// TIA Portal V18 export
FUNCTION "Interlock dos sinais linha" : Void   // FC9, LAD
{ S7_Optimized_Access := 'TRUE' }
// stored: SetENOAutomatically false
   VAR_TEMP
      SIGNAL_HELGE : Bool;
      SIGNAL_HELGE1 : Bool;
   END_VAR
   VAR_TEMP   // added for the SCL form of the ladder/FBD networks
      _w1 : Bool;
      _w2 : Bool;
      _w3 : Bool;
      _w4 : Bool;
   END_VAR
BEGIN

REGION Network 1: SCADA DESABILITADO
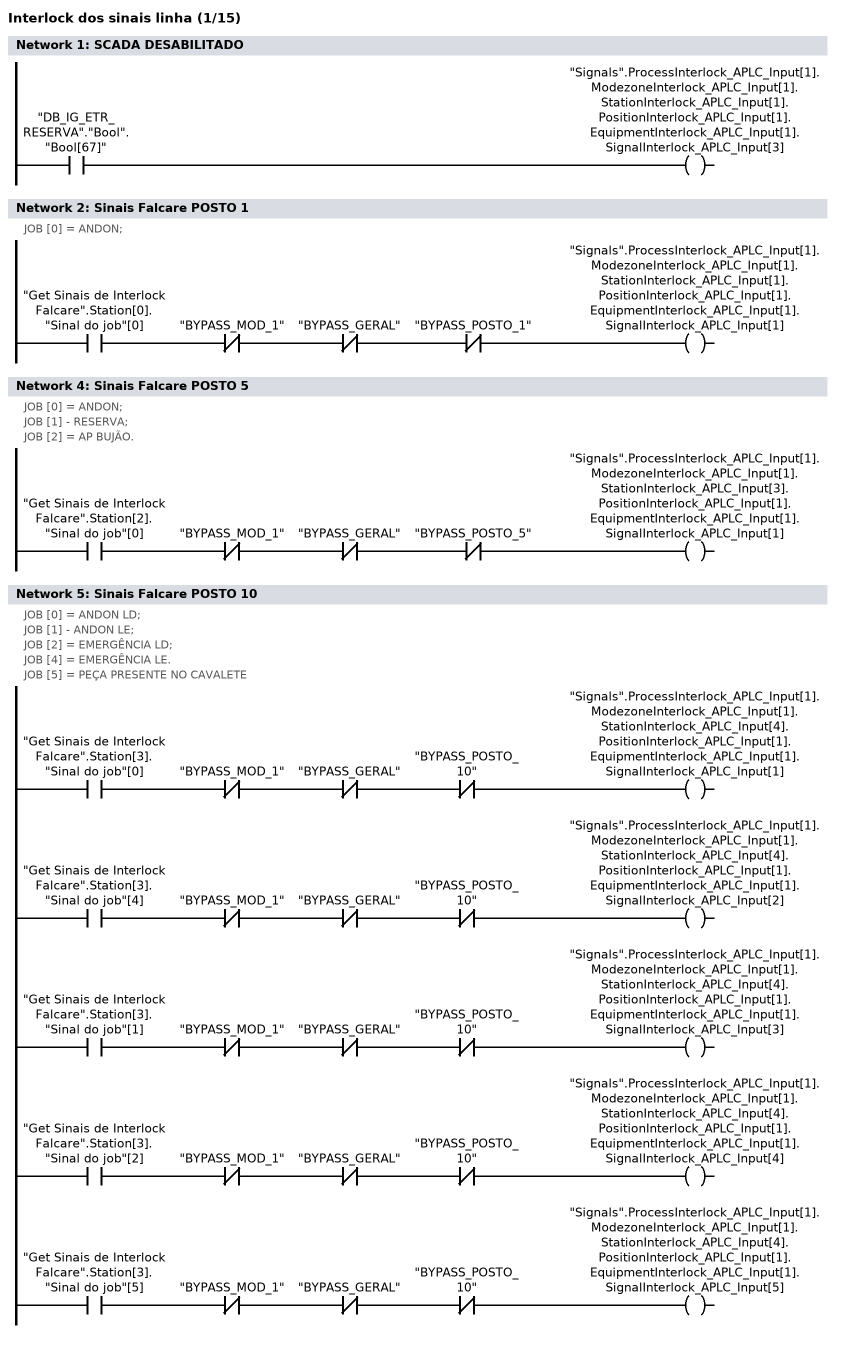
   RUNG wire#powerrail
      Contact( "DB_IG_ETR_RESERVA"."Bool"."Bool[67]" )
      Coil( "Signals".ProcessInterlock_APLC_Input[1].ModezoneInterlock_APLC_Input[1].StationInterlock_APLC_Input[1].PositionInterlock_APLC_Input[1].EquipmentInterlock_APLC_Input[1].SignalInterlock_APLC_Input[3] )
   END_RUNG
   // the same network as SCL:
   "Signals".ProcessInterlock_APLC_Input[1].ModezoneInterlock_APLC_Input[1].StationInterlock_APLC_Input[1].PositionInterlock_APLC_Input[1].EquipmentInterlock_APLC_Input[1].SignalInterlock_APLC_Input[3] := "DB_IG_ETR_RESERVA"."Bool"."Bool[67]";
END_REGION

REGION Network 2: Sinais Falcare POSTO 1
   // JOB [0] = ANDON;
   RUNG wire#powerrail
      Contact( "Get Sinais de Interlock Falcare".Station[0]."Sinal do job"[0] )
      I_Contact( "BYPASS_MOD_1" )
      I_Contact( "BYPASS_GERAL" )
      I_Contact( "BYPASS_POSTO_1" )
      Coil( "Signals".ProcessInterlock_APLC_Input[1].ModezoneInterlock_APLC_Input[1].StationInterlock_APLC_Input[1].PositionInterlock_APLC_Input[1].EquipmentInterlock_APLC_Input[1].SignalInterlock_APLC_Input[1] )
   END_RUNG
   // the same network as SCL:
   "Signals".ProcessInterlock_APLC_Input[1].ModezoneInterlock_APLC_Input[1].StationInterlock_APLC_Input[1].PositionInterlock_APLC_Input[1].EquipmentInterlock_APLC_Input[1].SignalInterlock_APLC_Input[1] := "Get Sinais de Interlock Falcare".Station[0]."Sinal do job"[0] AND NOT "BYPASS_MOD_1" AND NOT "BYPASS_GERAL" AND NOT "BYPASS_POSTO_1";
END_REGION

REGION Network 3: Sinais Falcare VIVERK
   // JOB [0] = ANDON;
   // JOB [1] - EMERGÊNCIA;
END_REGION

REGION Network 4: Sinais Falcare POSTO 5
   // JOB [0] = ANDON;
   // JOB [1] - RESERVA;
   // JOB [2] = AP BUJÃO.
   RUNG wire#powerrail
      Contact( "Get Sinais de Interlock Falcare".Station[2]."Sinal do job"[0] )
      I_Contact( "BYPASS_MOD_1" )
      I_Contact( "BYPASS_GERAL" )
      I_Contact( "BYPASS_POSTO_5" )
      Coil( "Signals".ProcessInterlock_APLC_Input[1].ModezoneInterlock_APLC_Input[1].StationInterlock_APLC_Input[3].PositionInterlock_APLC_Input[1].EquipmentInterlock_APLC_Input[1].SignalInterlock_APLC_Input[1] )
   END_RUNG
   // the same network as SCL:
   "Signals".ProcessInterlock_APLC_Input[1].ModezoneInterlock_APLC_Input[1].StationInterlock_APLC_Input[3].PositionInterlock_APLC_Input[1].EquipmentInterlock_APLC_Input[1].SignalInterlock_APLC_Input[1] := "Get Sinais de Interlock Falcare".Station[2]."Sinal do job"[0] AND NOT "BYPASS_MOD_1" AND NOT "BYPASS_GERAL" AND NOT "BYPASS_POSTO_5";
END_REGION

REGION Network 5: Sinais Falcare POSTO 10
   // JOB [0] = ANDON LD;
   // JOB [1] - ANDON LE;
   // JOB [2] = EMERGÊNCIA LD;
   // JOB [4] = EMERGÊNCIA LE.
   // JOB [5] = PEÇA PRESENTE NO CAVALETE
   RUNG wire#powerrail
      Contact( "Get Sinais de Interlock Falcare".Station[3]."Sinal do job"[0] )
      I_Contact( "BYPASS_MOD_1" )
      I_Contact( "BYPASS_GERAL" )
      I_Contact( "BYPASS_POSTO_10" )
      Coil( "Signals".ProcessInterlock_APLC_Input[1].ModezoneInterlock_APLC_Input[1].StationInterlock_APLC_Input[4].PositionInterlock_APLC_Input[1].EquipmentInterlock_APLC_Input[1].SignalInterlock_APLC_Input[1] )
   END_RUNG
   RUNG wire#powerrail
      Contact( "Get Sinais de Interlock Falcare".Station[3]."Sinal do job"[4] )
      I_Contact( "BYPASS_MOD_1" )
      I_Contact( "BYPASS_GERAL" )
      I_Contact( "BYPASS_POSTO_10" )
      Coil( "Signals".ProcessInterlock_APLC_Input[1].ModezoneInterlock_APLC_Input[1].StationInterlock_APLC_Input[4].PositionInterlock_APLC_Input[1].EquipmentInterlock_APLC_Input[1].SignalInterlock_APLC_Input[2] )
   END_RUNG
   RUNG wire#powerrail
      Contact( "Get Sinais de Interlock Falcare".Station[3]."Sinal do job"[1] )
      I_Contact( "BYPASS_MOD_1" )
      I_Contact( "BYPASS_GERAL" )
      I_Contact( "BYPASS_POSTO_10" )
      Coil( "Signals".ProcessInterlock_APLC_Input[1].ModezoneInterlock_APLC_Input[1].StationInterlock_APLC_Input[4].PositionInterlock_APLC_Input[1].EquipmentInterlock_APLC_Input[1].SignalInterlock_APLC_Input[3] )
   END_RUNG
   RUNG wire#powerrail
      Contact( "Get Sinais de Interlock Falcare".Station[3]."Sinal do job"[2] )
      I_Contact( "BYPASS_MOD_1" )
      I_Contact( "BYPASS_GERAL" )
      I_Contact( "BYPASS_POSTO_10" )
      Coil( "Signals".ProcessInterlock_APLC_Input[1].ModezoneInterlock_APLC_Input[1].StationInterlock_APLC_Input[4].PositionInterlock_APLC_Input[1].EquipmentInterlock_APLC_Input[1].SignalInterlock_APLC_Input[4] )
   END_RUNG
   RUNG wire#powerrail
      Contact( "Get Sinais de Interlock Falcare".Station[3]."Sinal do job"[5] )
      I_Contact( "BYPASS_MOD_1" )
      I_Contact( "BYPASS_GERAL" )
      I_Contact( "BYPASS_POSTO_10" )
      Coil( "Signals".ProcessInterlock_APLC_Input[1].ModezoneInterlock_APLC_Input[1].StationInterlock_APLC_Input[4].PositionInterlock_APLC_Input[1].EquipmentInterlock_APLC_Input[1].SignalInterlock_APLC_Input[5] )
   END_RUNG
   // the same network as SCL:
   "Signals".ProcessInterlock_APLC_Input[1].ModezoneInterlock_APLC_Input[1].StationInterlock_APLC_Input[4].PositionInterlock_APLC_Input[1].EquipmentInterlock_APLC_Input[1].SignalInterlock_APLC_Input[1] := "Get Sinais de Interlock Falcare".Station[3]."Sinal do job"[0] AND NOT "BYPASS_MOD_1" AND NOT "BYPASS_GERAL" AND NOT "BYPASS_POSTO_10";
   "Signals".ProcessInterlock_APLC_Input[1].ModezoneInterlock_APLC_Input[1].StationInterlock_APLC_Input[4].PositionInterlock_APLC_Input[1].EquipmentInterlock_APLC_Input[1].SignalInterlock_APLC_Input[2] := "Get Sinais de Interlock Falcare".Station[3]."Sinal do job"[4] AND NOT "BYPASS_MOD_1" AND NOT "BYPASS_GERAL" AND NOT "BYPASS_POSTO_10";
   "Signals".ProcessInterlock_APLC_Input[1].ModezoneInterlock_APLC_Input[1].StationInterlock_APLC_Input[4].PositionInterlock_APLC_Input[1].EquipmentInterlock_APLC_Input[1].SignalInterlock_APLC_Input[3] := "Get Sinais de Interlock Falcare".Station[3]."Sinal do job"[1] AND NOT "BYPASS_MOD_1" AND NOT "BYPASS_GERAL" AND NOT "BYPASS_POSTO_10";
   "Signals".ProcessInterlock_APLC_Input[1].ModezoneInterlock_APLC_Input[1].StationInterlock_APLC_Input[4].PositionInterlock_APLC_Input[1].EquipmentInterlock_APLC_Input[1].SignalInterlock_APLC_Input[4] := "Get Sinais de Interlock Falcare".Station[3]."Sinal do job"[2] AND NOT "BYPASS_MOD_1" AND NOT "BYPASS_GERAL" AND NOT "BYPASS_POSTO_10";
   "Signals".ProcessInterlock_APLC_Input[1].ModezoneInterlock_APLC_Input[1].StationInterlock_APLC_Input[4].PositionInterlock_APLC_Input[1].EquipmentInterlock_APLC_Input[1].SignalInterlock_APLC_Input[5] := "Get Sinais de Interlock Falcare".Station[3]."Sinal do job"[5] AND NOT "BYPASS_MOD_1" AND NOT "BYPASS_GERAL" AND NOT "BYPASS_POSTO_10";
END_REGION

REGION Network 6: Sinais Falcare POSTO 15
   // JOB [3] = AP TUBO RPX POSTO 15;
END_REGION

REGION Network 7: Sinais Falcare POSTO 20
   // JOB [0] = ANDON LD;
   // JOB [1] - EMERGÊNCIA LD;
   // JOB [2] = AP MOLA HARPA;
   // JOB [3] = SENSOR POSIÇÃO AP HARPA;
   // JOB [4] = AP TUBO LUBRIFICAÇÃO RPX I9.0
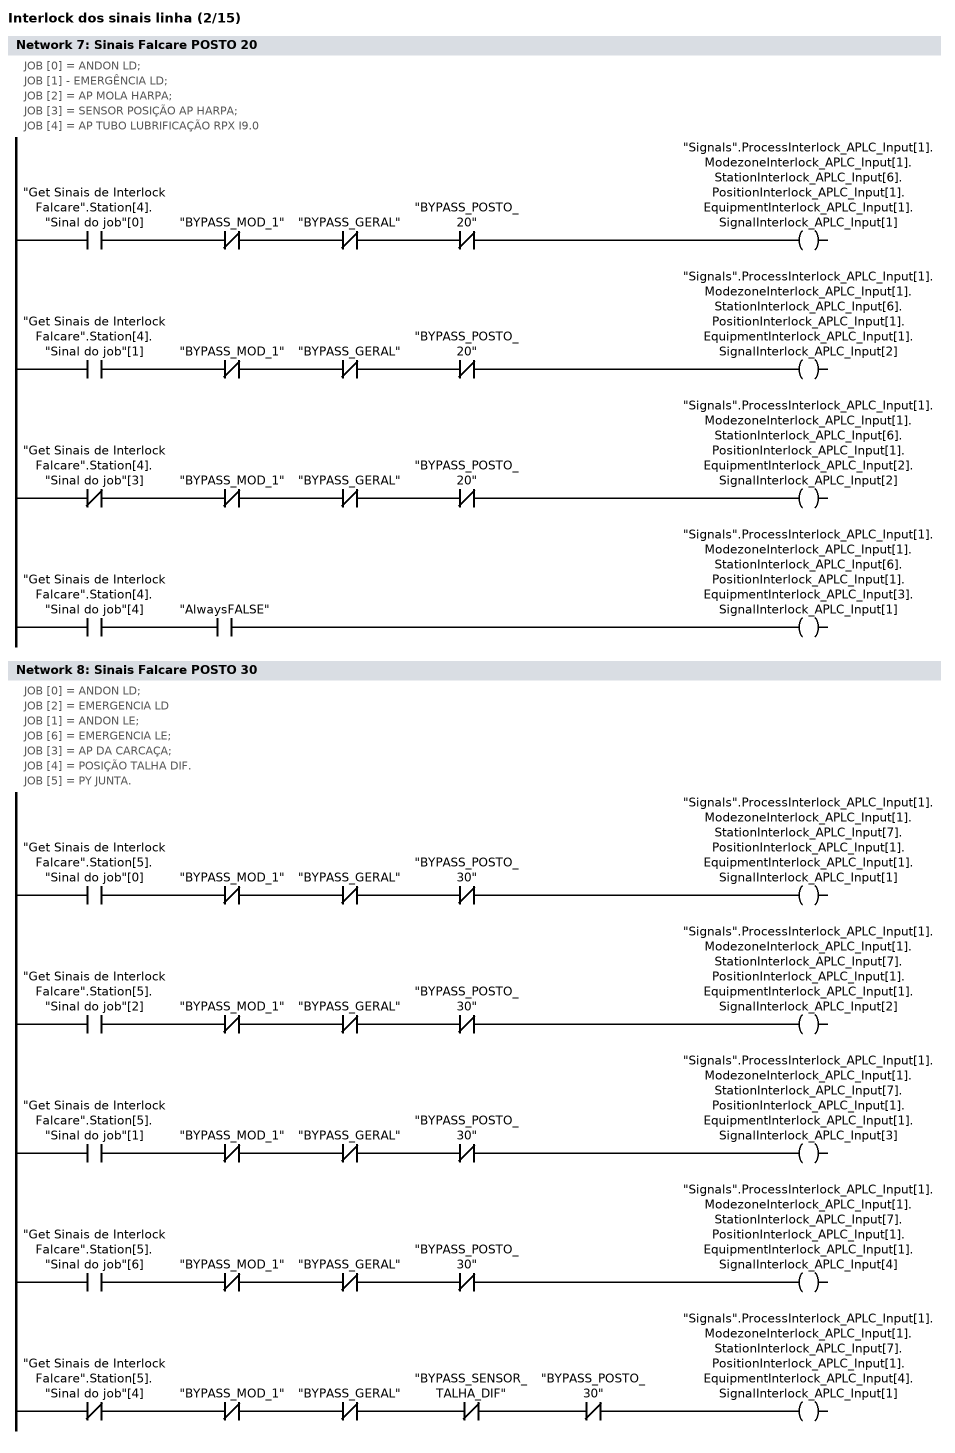
   RUNG wire#powerrail
      Contact( "Get Sinais de Interlock Falcare".Station[4]."Sinal do job"[0] )
      I_Contact( "BYPASS_MOD_1" )
      I_Contact( "BYPASS_GERAL" )
      I_Contact( "BYPASS_POSTO_20" )
      Coil( "Signals".ProcessInterlock_APLC_Input[1].ModezoneInterlock_APLC_Input[1].StationInterlock_APLC_Input[6].PositionInterlock_APLC_Input[1].EquipmentInterlock_APLC_Input[1].SignalInterlock_APLC_Input[1] )
   END_RUNG
   RUNG wire#powerrail
      Contact( "Get Sinais de Interlock Falcare".Station[4]."Sinal do job"[1] )
      I_Contact( "BYPASS_MOD_1" )
      I_Contact( "BYPASS_GERAL" )
      I_Contact( "BYPASS_POSTO_20" )
      Coil( "Signals".ProcessInterlock_APLC_Input[1].ModezoneInterlock_APLC_Input[1].StationInterlock_APLC_Input[6].PositionInterlock_APLC_Input[1].EquipmentInterlock_APLC_Input[1].SignalInterlock_APLC_Input[2] )
   END_RUNG
   RUNG wire#powerrail
      I_Contact( "Get Sinais de Interlock Falcare".Station[4]."Sinal do job"[3] )
      I_Contact( "BYPASS_MOD_1" )
      I_Contact( "BYPASS_GERAL" )
      I_Contact( "BYPASS_POSTO_20" )
      Coil( "Signals".ProcessInterlock_APLC_Input[1].ModezoneInterlock_APLC_Input[1].StationInterlock_APLC_Input[6].PositionInterlock_APLC_Input[1].EquipmentInterlock_APLC_Input[2].SignalInterlock_APLC_Input[2] )
   END_RUNG
   RUNG wire#powerrail
      Contact( "Get Sinais de Interlock Falcare".Station[4]."Sinal do job"[4] )
      Contact( "AlwaysFALSE" )
      Coil( "Signals".ProcessInterlock_APLC_Input[1].ModezoneInterlock_APLC_Input[1].StationInterlock_APLC_Input[6].PositionInterlock_APLC_Input[1].EquipmentInterlock_APLC_Input[3].SignalInterlock_APLC_Input[1] )
   END_RUNG
   // the same network as SCL:
   "Signals".ProcessInterlock_APLC_Input[1].ModezoneInterlock_APLC_Input[1].StationInterlock_APLC_Input[6].PositionInterlock_APLC_Input[1].EquipmentInterlock_APLC_Input[1].SignalInterlock_APLC_Input[1] := "Get Sinais de Interlock Falcare".Station[4]."Sinal do job"[0] AND NOT "BYPASS_MOD_1" AND NOT "BYPASS_GERAL" AND NOT "BYPASS_POSTO_20";
   "Signals".ProcessInterlock_APLC_Input[1].ModezoneInterlock_APLC_Input[1].StationInterlock_APLC_Input[6].PositionInterlock_APLC_Input[1].EquipmentInterlock_APLC_Input[1].SignalInterlock_APLC_Input[2] := "Get Sinais de Interlock Falcare".Station[4]."Sinal do job"[1] AND NOT "BYPASS_MOD_1" AND NOT "BYPASS_GERAL" AND NOT "BYPASS_POSTO_20";
   "Signals".ProcessInterlock_APLC_Input[1].ModezoneInterlock_APLC_Input[1].StationInterlock_APLC_Input[6].PositionInterlock_APLC_Input[1].EquipmentInterlock_APLC_Input[2].SignalInterlock_APLC_Input[2] := NOT "Get Sinais de Interlock Falcare".Station[4]."Sinal do job"[3] AND NOT "BYPASS_MOD_1" AND NOT "BYPASS_GERAL" AND NOT "BYPASS_POSTO_20";
   "Signals".ProcessInterlock_APLC_Input[1].ModezoneInterlock_APLC_Input[1].StationInterlock_APLC_Input[6].PositionInterlock_APLC_Input[1].EquipmentInterlock_APLC_Input[3].SignalInterlock_APLC_Input[1] := "Get Sinais de Interlock Falcare".Station[4]."Sinal do job"[4] AND "AlwaysFALSE";
END_REGION

REGION Network 8: Sinais Falcare POSTO 30
   // JOB [0] = ANDON LD;
   // JOB [2] = EMERGENCIA LD
   // JOB [1] = ANDON LE;
   // JOB [6] = EMERGENCIA LE;
   // JOB [3] = AP DA CARCAÇA;
   // JOB [4] = POSIÇÃO TALHA DIF.
   // JOB [5] = PY JUNTA.
   RUNG wire#powerrail
      Contact( "Get Sinais de Interlock Falcare".Station[5]."Sinal do job"[0] )
      I_Contact( "BYPASS_MOD_1" )
      I_Contact( "BYPASS_GERAL" )
      I_Contact( "BYPASS_POSTO_30" )
      Coil( "Signals".ProcessInterlock_APLC_Input[1].ModezoneInterlock_APLC_Input[1].StationInterlock_APLC_Input[7].PositionInterlock_APLC_Input[1].EquipmentInterlock_APLC_Input[1].SignalInterlock_APLC_Input[1] )
   END_RUNG
   RUNG wire#powerrail
      Contact( "Get Sinais de Interlock Falcare".Station[5]."Sinal do job"[2] )
      I_Contact( "BYPASS_MOD_1" )
      I_Contact( "BYPASS_GERAL" )
      I_Contact( "BYPASS_POSTO_30" )
      Coil( "Signals".ProcessInterlock_APLC_Input[1].ModezoneInterlock_APLC_Input[1].StationInterlock_APLC_Input[7].PositionInterlock_APLC_Input[1].EquipmentInterlock_APLC_Input[1].SignalInterlock_APLC_Input[2] )
   END_RUNG
   RUNG wire#powerrail
      Contact( "Get Sinais de Interlock Falcare".Station[5]."Sinal do job"[1] )
      I_Contact( "BYPASS_MOD_1" )
      I_Contact( "BYPASS_GERAL" )
      I_Contact( "BYPASS_POSTO_30" )
      Coil( "Signals".ProcessInterlock_APLC_Input[1].ModezoneInterlock_APLC_Input[1].StationInterlock_APLC_Input[7].PositionInterlock_APLC_Input[1].EquipmentInterlock_APLC_Input[1].SignalInterlock_APLC_Input[3] )
   END_RUNG
   RUNG wire#powerrail
      Contact( "Get Sinais de Interlock Falcare".Station[5]."Sinal do job"[6] )
      I_Contact( "BYPASS_MOD_1" )
      I_Contact( "BYPASS_GERAL" )
      I_Contact( "BYPASS_POSTO_30" )
      Coil( "Signals".ProcessInterlock_APLC_Input[1].ModezoneInterlock_APLC_Input[1].StationInterlock_APLC_Input[7].PositionInterlock_APLC_Input[1].EquipmentInterlock_APLC_Input[1].SignalInterlock_APLC_Input[4] )
   END_RUNG
   RUNG wire#powerrail
      I_Contact( "Get Sinais de Interlock Falcare".Station[5]."Sinal do job"[4] )
      I_Contact( "BYPASS_MOD_1" )
      I_Contact( "BYPASS_GERAL" )
      I_Contact( "BYPASS_SENSOR_TALHA_DIF" )
      I_Contact( "BYPASS_POSTO_30" )
      Coil( "Signals".ProcessInterlock_APLC_Input[1].ModezoneInterlock_APLC_Input[1].StationInterlock_APLC_Input[7].PositionInterlock_APLC_Input[1].EquipmentInterlock_APLC_Input[4].SignalInterlock_APLC_Input[1] )
   END_RUNG
   // the same network as SCL:
   "Signals".ProcessInterlock_APLC_Input[1].ModezoneInterlock_APLC_Input[1].StationInterlock_APLC_Input[7].PositionInterlock_APLC_Input[1].EquipmentInterlock_APLC_Input[1].SignalInterlock_APLC_Input[1] := "Get Sinais de Interlock Falcare".Station[5]."Sinal do job"[0] AND NOT "BYPASS_MOD_1" AND NOT "BYPASS_GERAL" AND NOT "BYPASS_POSTO_30";
   "Signals".ProcessInterlock_APLC_Input[1].ModezoneInterlock_APLC_Input[1].StationInterlock_APLC_Input[7].PositionInterlock_APLC_Input[1].EquipmentInterlock_APLC_Input[1].SignalInterlock_APLC_Input[2] := "Get Sinais de Interlock Falcare".Station[5]."Sinal do job"[2] AND NOT "BYPASS_MOD_1" AND NOT "BYPASS_GERAL" AND NOT "BYPASS_POSTO_30";
   "Signals".ProcessInterlock_APLC_Input[1].ModezoneInterlock_APLC_Input[1].StationInterlock_APLC_Input[7].PositionInterlock_APLC_Input[1].EquipmentInterlock_APLC_Input[1].SignalInterlock_APLC_Input[3] := "Get Sinais de Interlock Falcare".Station[5]."Sinal do job"[1] AND NOT "BYPASS_MOD_1" AND NOT "BYPASS_GERAL" AND NOT "BYPASS_POSTO_30";
   "Signals".ProcessInterlock_APLC_Input[1].ModezoneInterlock_APLC_Input[1].StationInterlock_APLC_Input[7].PositionInterlock_APLC_Input[1].EquipmentInterlock_APLC_Input[1].SignalInterlock_APLC_Input[4] := "Get Sinais de Interlock Falcare".Station[5]."Sinal do job"[6] AND NOT "BYPASS_MOD_1" AND NOT "BYPASS_GERAL" AND NOT "BYPASS_POSTO_30";
   "Signals".ProcessInterlock_APLC_Input[1].ModezoneInterlock_APLC_Input[1].StationInterlock_APLC_Input[7].PositionInterlock_APLC_Input[1].EquipmentInterlock_APLC_Input[4].SignalInterlock_APLC_Input[1] := NOT "Get Sinais de Interlock Falcare".Station[5]."Sinal do job"[4] AND NOT "BYPASS_MOD_1" AND NOT "BYPASS_GERAL" AND NOT "BYPASS_SENSOR_TALHA_DIF" AND NOT "BYPASS_POSTO_30";
END_REGION

REGION Network 9: Sinais Falcare POSTO 40
   // JOB [0] = ANDON LD;
   // JOB [1] = ANDON LE;
   // JOB [2] = EMERGENCIA LE;
   // JOB [3] = AP CRAWFOOT PORCA;
   // JOB [4] = SENSOR POSIÇÃO AP CRAWFOOT;
   // JOB [5] = AP PORCA DUPLO FUSO;
   // JOB [6] = SENSOR POSIÇÃO AP DUPLO FUSO;
   // JOB [7] = EMERGÊNCIA LD.
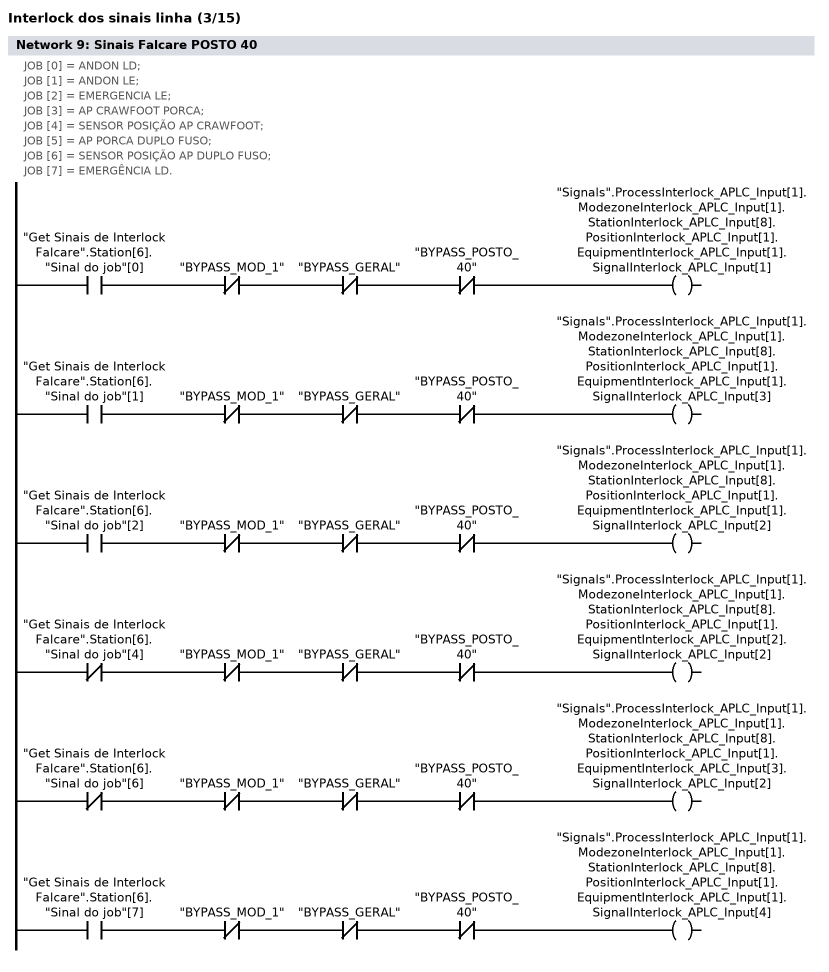
   RUNG wire#powerrail
      Contact( "Get Sinais de Interlock Falcare".Station[6]."Sinal do job"[0] )
      I_Contact( "BYPASS_MOD_1" )
      I_Contact( "BYPASS_GERAL" )
      I_Contact( "BYPASS_POSTO_40" )
      Coil( "Signals".ProcessInterlock_APLC_Input[1].ModezoneInterlock_APLC_Input[1].StationInterlock_APLC_Input[8].PositionInterlock_APLC_Input[1].EquipmentInterlock_APLC_Input[1].SignalInterlock_APLC_Input[1] )
   END_RUNG
   RUNG wire#powerrail
      Contact( "Get Sinais de Interlock Falcare".Station[6]."Sinal do job"[1] )
      I_Contact( "BYPASS_MOD_1" )
      I_Contact( "BYPASS_GERAL" )
      I_Contact( "BYPASS_POSTO_40" )
      Coil( "Signals".ProcessInterlock_APLC_Input[1].ModezoneInterlock_APLC_Input[1].StationInterlock_APLC_Input[8].PositionInterlock_APLC_Input[1].EquipmentInterlock_APLC_Input[1].SignalInterlock_APLC_Input[3] )
   END_RUNG
   RUNG wire#powerrail
      Contact( "Get Sinais de Interlock Falcare".Station[6]."Sinal do job"[2] )
      I_Contact( "BYPASS_MOD_1" )
      I_Contact( "BYPASS_GERAL" )
      I_Contact( "BYPASS_POSTO_40" )
      Coil( "Signals".ProcessInterlock_APLC_Input[1].ModezoneInterlock_APLC_Input[1].StationInterlock_APLC_Input[8].PositionInterlock_APLC_Input[1].EquipmentInterlock_APLC_Input[1].SignalInterlock_APLC_Input[2] )
   END_RUNG
   RUNG wire#powerrail
      I_Contact( "Get Sinais de Interlock Falcare".Station[6]."Sinal do job"[4] )
      I_Contact( "BYPASS_MOD_1" )
      I_Contact( "BYPASS_GERAL" )
      I_Contact( "BYPASS_POSTO_40" )
      Coil( "Signals".ProcessInterlock_APLC_Input[1].ModezoneInterlock_APLC_Input[1].StationInterlock_APLC_Input[8].PositionInterlock_APLC_Input[1].EquipmentInterlock_APLC_Input[2].SignalInterlock_APLC_Input[2] )
   END_RUNG
   RUNG wire#powerrail
      I_Contact( "Get Sinais de Interlock Falcare".Station[6]."Sinal do job"[6] )
      I_Contact( "BYPASS_MOD_1" )
      I_Contact( "BYPASS_GERAL" )
      I_Contact( "BYPASS_POSTO_40" )
      Coil( "Signals".ProcessInterlock_APLC_Input[1].ModezoneInterlock_APLC_Input[1].StationInterlock_APLC_Input[8].PositionInterlock_APLC_Input[1].EquipmentInterlock_APLC_Input[3].SignalInterlock_APLC_Input[2] )
   END_RUNG
   RUNG wire#powerrail
      Contact( "Get Sinais de Interlock Falcare".Station[6]."Sinal do job"[7] )
      I_Contact( "BYPASS_MOD_1" )
      I_Contact( "BYPASS_GERAL" )
      I_Contact( "BYPASS_POSTO_40" )
      Coil( "Signals".ProcessInterlock_APLC_Input[1].ModezoneInterlock_APLC_Input[1].StationInterlock_APLC_Input[8].PositionInterlock_APLC_Input[1].EquipmentInterlock_APLC_Input[1].SignalInterlock_APLC_Input[4] )
   END_RUNG
   // the same network as SCL:
   "Signals".ProcessInterlock_APLC_Input[1].ModezoneInterlock_APLC_Input[1].StationInterlock_APLC_Input[8].PositionInterlock_APLC_Input[1].EquipmentInterlock_APLC_Input[1].SignalInterlock_APLC_Input[1] := "Get Sinais de Interlock Falcare".Station[6]."Sinal do job"[0] AND NOT "BYPASS_MOD_1" AND NOT "BYPASS_GERAL" AND NOT "BYPASS_POSTO_40";
   "Signals".ProcessInterlock_APLC_Input[1].ModezoneInterlock_APLC_Input[1].StationInterlock_APLC_Input[8].PositionInterlock_APLC_Input[1].EquipmentInterlock_APLC_Input[1].SignalInterlock_APLC_Input[3] := "Get Sinais de Interlock Falcare".Station[6]."Sinal do job"[1] AND NOT "BYPASS_MOD_1" AND NOT "BYPASS_GERAL" AND NOT "BYPASS_POSTO_40";
   "Signals".ProcessInterlock_APLC_Input[1].ModezoneInterlock_APLC_Input[1].StationInterlock_APLC_Input[8].PositionInterlock_APLC_Input[1].EquipmentInterlock_APLC_Input[1].SignalInterlock_APLC_Input[2] := "Get Sinais de Interlock Falcare".Station[6]."Sinal do job"[2] AND NOT "BYPASS_MOD_1" AND NOT "BYPASS_GERAL" AND NOT "BYPASS_POSTO_40";
   "Signals".ProcessInterlock_APLC_Input[1].ModezoneInterlock_APLC_Input[1].StationInterlock_APLC_Input[8].PositionInterlock_APLC_Input[1].EquipmentInterlock_APLC_Input[2].SignalInterlock_APLC_Input[2] := NOT "Get Sinais de Interlock Falcare".Station[6]."Sinal do job"[4] AND NOT "BYPASS_MOD_1" AND NOT "BYPASS_GERAL" AND NOT "BYPASS_POSTO_40";
   "Signals".ProcessInterlock_APLC_Input[1].ModezoneInterlock_APLC_Input[1].StationInterlock_APLC_Input[8].PositionInterlock_APLC_Input[1].EquipmentInterlock_APLC_Input[3].SignalInterlock_APLC_Input[2] := NOT "Get Sinais de Interlock Falcare".Station[6]."Sinal do job"[6] AND NOT "BYPASS_MOD_1" AND NOT "BYPASS_GERAL" AND NOT "BYPASS_POSTO_40";
   "Signals".ProcessInterlock_APLC_Input[1].ModezoneInterlock_APLC_Input[1].StationInterlock_APLC_Input[8].PositionInterlock_APLC_Input[1].EquipmentInterlock_APLC_Input[1].SignalInterlock_APLC_Input[4] := "Get Sinais de Interlock Falcare".Station[6]."Sinal do job"[7] AND NOT "BYPASS_MOD_1" AND NOT "BYPASS_GERAL" AND NOT "BYPASS_POSTO_40";
END_REGION

REGION Network 10: Sinais Falcare POSTO 50
   // JOB [0] = ANDON;
   // JOB [1] = EMERGENCIA;
   // JOB [2] = AP PORCA ESCONDIDA;
   // JOB [3] = SENSOR POSIÇÃO AP PORCA ESCONDIDA;
   // JOB [4] = AP PORCA SUPORTE DO CILINDRO;
   // JOB [5] = SENSOR POSIÇÃO AP SUPORTE DO CILINDRO;
   // JOB [7] = AP VÁLVULA
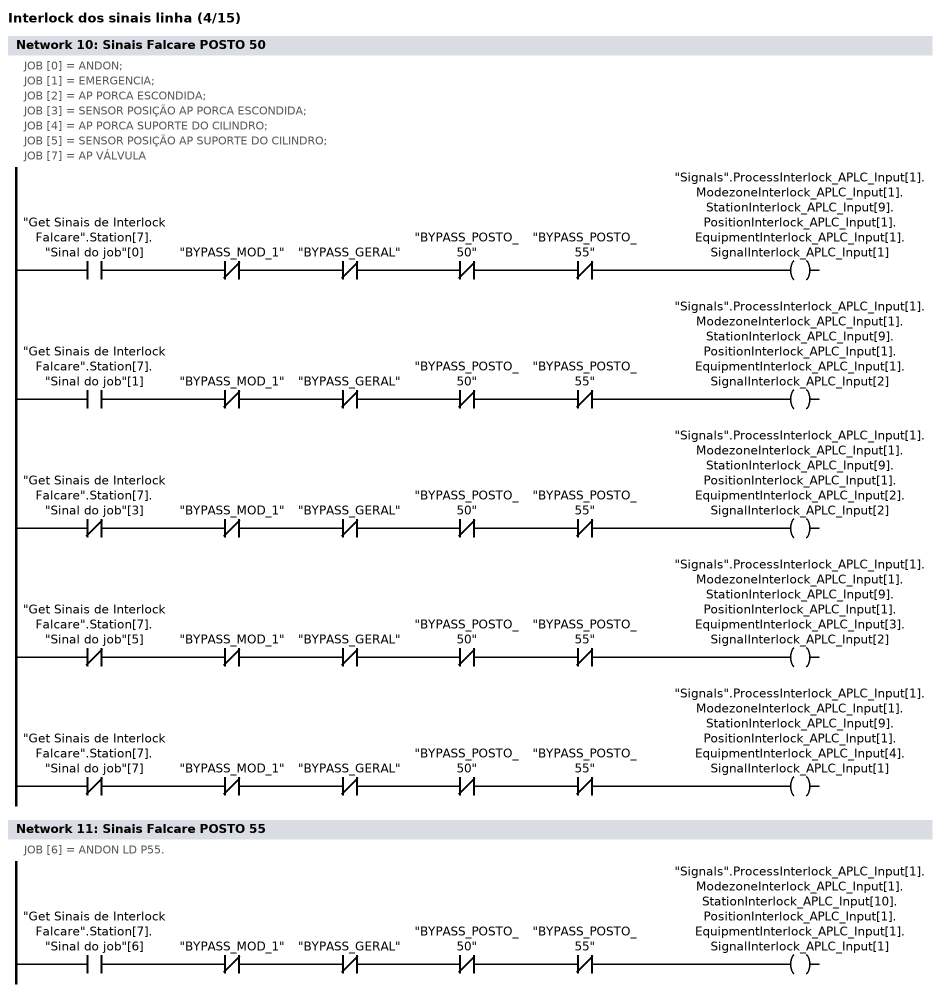
   RUNG wire#powerrail
      Contact( "Get Sinais de Interlock Falcare".Station[7]."Sinal do job"[0] )
      I_Contact( "BYPASS_MOD_1" )
      I_Contact( "BYPASS_GERAL" )
      I_Contact( "BYPASS_POSTO_50" )
      I_Contact( "BYPASS_POSTO_55" )
      Coil( "Signals".ProcessInterlock_APLC_Input[1].ModezoneInterlock_APLC_Input[1].StationInterlock_APLC_Input[9].PositionInterlock_APLC_Input[1].EquipmentInterlock_APLC_Input[1].SignalInterlock_APLC_Input[1] )
   END_RUNG
   RUNG wire#powerrail
      Contact( "Get Sinais de Interlock Falcare".Station[7]."Sinal do job"[1] )
      I_Contact( "BYPASS_MOD_1" )
      I_Contact( "BYPASS_GERAL" )
      I_Contact( "BYPASS_POSTO_50" )
      I_Contact( "BYPASS_POSTO_55" )
      Coil( "Signals".ProcessInterlock_APLC_Input[1].ModezoneInterlock_APLC_Input[1].StationInterlock_APLC_Input[9].PositionInterlock_APLC_Input[1].EquipmentInterlock_APLC_Input[1].SignalInterlock_APLC_Input[2] )
   END_RUNG
   RUNG wire#powerrail
      I_Contact( "Get Sinais de Interlock Falcare".Station[7]."Sinal do job"[3] )
      I_Contact( "BYPASS_MOD_1" )
      I_Contact( "BYPASS_GERAL" )
      I_Contact( "BYPASS_POSTO_50" )
      I_Contact( "BYPASS_POSTO_55" )
      Coil( "Signals".ProcessInterlock_APLC_Input[1].ModezoneInterlock_APLC_Input[1].StationInterlock_APLC_Input[9].PositionInterlock_APLC_Input[1].EquipmentInterlock_APLC_Input[2].SignalInterlock_APLC_Input[2] )
   END_RUNG
   RUNG wire#powerrail
      I_Contact( "Get Sinais de Interlock Falcare".Station[7]."Sinal do job"[5] )
      I_Contact( "BYPASS_MOD_1" )
      I_Contact( "BYPASS_GERAL" )
      I_Contact( "BYPASS_POSTO_50" )
      I_Contact( "BYPASS_POSTO_55" )
      Coil( "Signals".ProcessInterlock_APLC_Input[1].ModezoneInterlock_APLC_Input[1].StationInterlock_APLC_Input[9].PositionInterlock_APLC_Input[1].EquipmentInterlock_APLC_Input[3].SignalInterlock_APLC_Input[2] )
   END_RUNG
   RUNG wire#powerrail
      I_Contact( "Get Sinais de Interlock Falcare".Station[7]."Sinal do job"[7] )
      I_Contact( "BYPASS_MOD_1" )
      I_Contact( "BYPASS_GERAL" )
      I_Contact( "BYPASS_POSTO_50" )
      I_Contact( "BYPASS_POSTO_55" )
      Coil( "Signals".ProcessInterlock_APLC_Input[1].ModezoneInterlock_APLC_Input[1].StationInterlock_APLC_Input[9].PositionInterlock_APLC_Input[1].EquipmentInterlock_APLC_Input[4].SignalInterlock_APLC_Input[1] )
   END_RUNG
   // the same network as SCL:
   "Signals".ProcessInterlock_APLC_Input[1].ModezoneInterlock_APLC_Input[1].StationInterlock_APLC_Input[9].PositionInterlock_APLC_Input[1].EquipmentInterlock_APLC_Input[1].SignalInterlock_APLC_Input[1] := "Get Sinais de Interlock Falcare".Station[7]."Sinal do job"[0] AND NOT "BYPASS_MOD_1" AND NOT "BYPASS_GERAL" AND NOT "BYPASS_POSTO_50" AND NOT "BYPASS_POSTO_55";
   "Signals".ProcessInterlock_APLC_Input[1].ModezoneInterlock_APLC_Input[1].StationInterlock_APLC_Input[9].PositionInterlock_APLC_Input[1].EquipmentInterlock_APLC_Input[1].SignalInterlock_APLC_Input[2] := "Get Sinais de Interlock Falcare".Station[7]."Sinal do job"[1] AND NOT "BYPASS_MOD_1" AND NOT "BYPASS_GERAL" AND NOT "BYPASS_POSTO_50" AND NOT "BYPASS_POSTO_55";
   "Signals".ProcessInterlock_APLC_Input[1].ModezoneInterlock_APLC_Input[1].StationInterlock_APLC_Input[9].PositionInterlock_APLC_Input[1].EquipmentInterlock_APLC_Input[2].SignalInterlock_APLC_Input[2] := NOT "Get Sinais de Interlock Falcare".Station[7]."Sinal do job"[3] AND NOT "BYPASS_MOD_1" AND NOT "BYPASS_GERAL" AND NOT "BYPASS_POSTO_50" AND NOT "BYPASS_POSTO_55";
   "Signals".ProcessInterlock_APLC_Input[1].ModezoneInterlock_APLC_Input[1].StationInterlock_APLC_Input[9].PositionInterlock_APLC_Input[1].EquipmentInterlock_APLC_Input[3].SignalInterlock_APLC_Input[2] := NOT "Get Sinais de Interlock Falcare".Station[7]."Sinal do job"[5] AND NOT "BYPASS_MOD_1" AND NOT "BYPASS_GERAL" AND NOT "BYPASS_POSTO_50" AND NOT "BYPASS_POSTO_55";
   "Signals".ProcessInterlock_APLC_Input[1].ModezoneInterlock_APLC_Input[1].StationInterlock_APLC_Input[9].PositionInterlock_APLC_Input[1].EquipmentInterlock_APLC_Input[4].SignalInterlock_APLC_Input[1] := NOT "Get Sinais de Interlock Falcare".Station[7]."Sinal do job"[7] AND NOT "BYPASS_MOD_1" AND NOT "BYPASS_GERAL" AND NOT "BYPASS_POSTO_50" AND NOT "BYPASS_POSTO_55";
END_REGION

REGION Network 11: Sinais Falcare POSTO 55
   // JOB [6] = ANDON LD P55.
   RUNG wire#powerrail
      Contact( "Get Sinais de Interlock Falcare".Station[7]."Sinal do job"[6] )
      I_Contact( "BYPASS_MOD_1" )
      I_Contact( "BYPASS_GERAL" )
      I_Contact( "BYPASS_POSTO_50" )
      I_Contact( "BYPASS_POSTO_55" )
      Coil( "Signals".ProcessInterlock_APLC_Input[1].ModezoneInterlock_APLC_Input[1].StationInterlock_APLC_Input[10].PositionInterlock_APLC_Input[1].EquipmentInterlock_APLC_Input[1].SignalInterlock_APLC_Input[1] )
   END_RUNG
   // the same network as SCL:
   "Signals".ProcessInterlock_APLC_Input[1].ModezoneInterlock_APLC_Input[1].StationInterlock_APLC_Input[10].PositionInterlock_APLC_Input[1].EquipmentInterlock_APLC_Input[1].SignalInterlock_APLC_Input[1] := "Get Sinais de Interlock Falcare".Station[7]."Sinal do job"[6] AND NOT "BYPASS_MOD_1" AND NOT "BYPASS_GERAL" AND NOT "BYPASS_POSTO_50" AND NOT "BYPASS_POSTO_55";
END_REGION

REGION Network 12: Sinais Falcare POSTO 60
   // JOB [0] = ANDON;
   // JOB [1] = EMERGENCIA;
   // JOB [2] = AP PORCA DO CILINDRO;
   // JOB [3] = SENSOR POSIÇÃO AP PORCA DO CILINDRO;
   // JOB [4] = EMERGENCIA PAINEL FALCARE.
   // JOB [5] = CONFIRMA PRE AVISO DO GIRADOR
   // JOB [6] = PRODUTO PRESENTE NO GIRADOR (MENSAGEM DE RETIRAR PRODUTO)
   // JOB [7] = FALCARE EM MANUAL
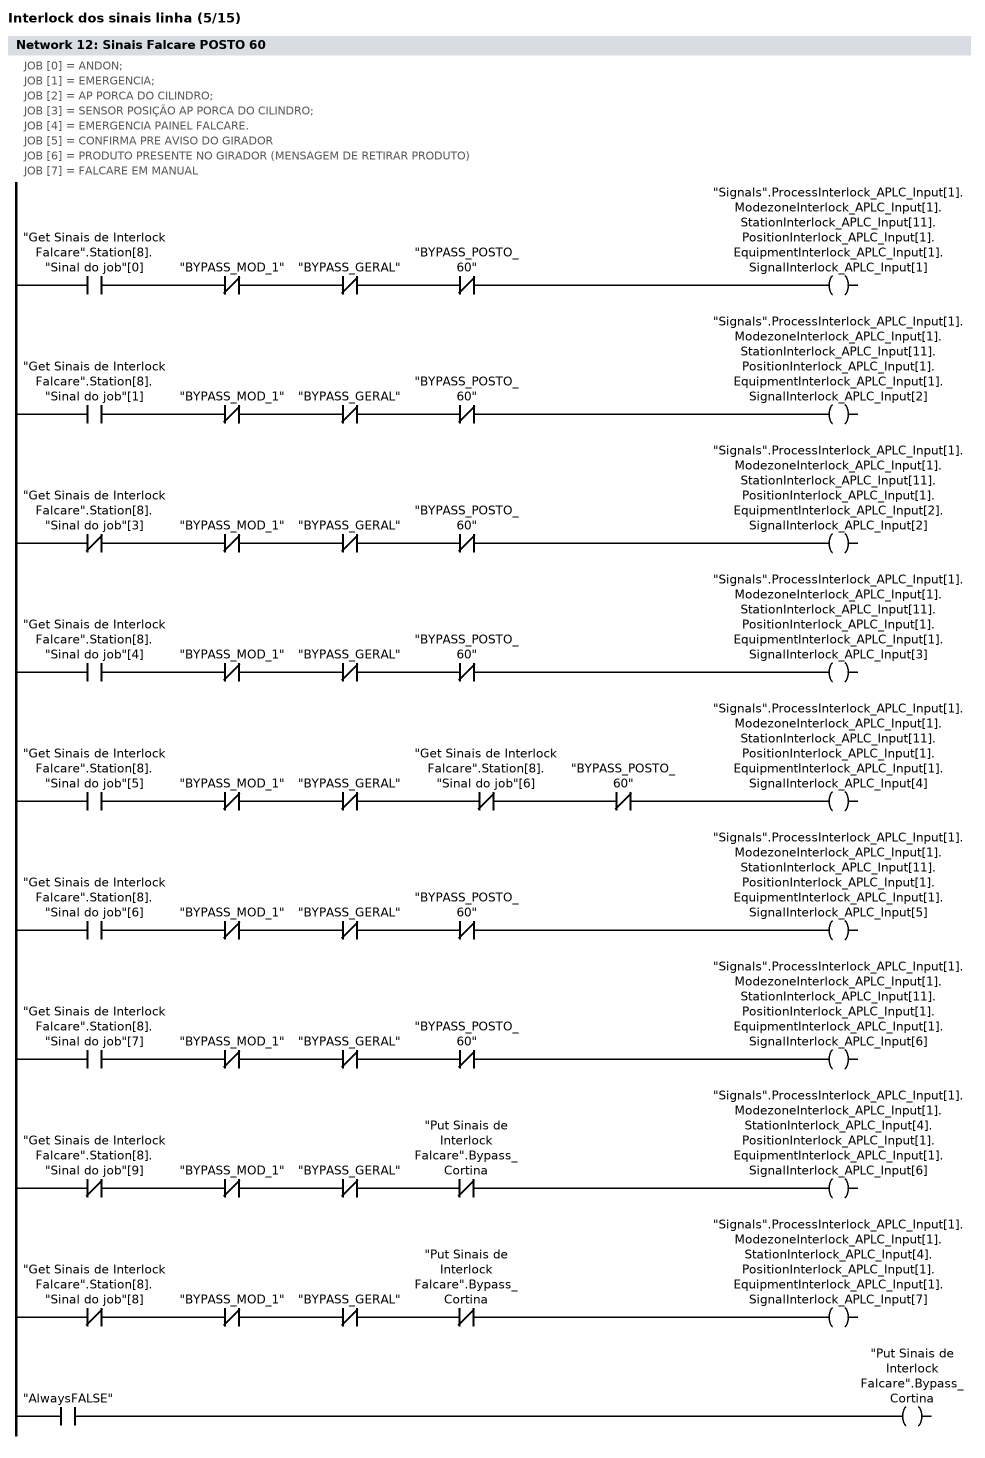
   RUNG wire#powerrail
      Contact( "Get Sinais de Interlock Falcare".Station[8]."Sinal do job"[0] )
      I_Contact( "BYPASS_MOD_1" )
      I_Contact( "BYPASS_GERAL" )
      I_Contact( "BYPASS_POSTO_60" )
      Coil( "Signals".ProcessInterlock_APLC_Input[1].ModezoneInterlock_APLC_Input[1].StationInterlock_APLC_Input[11].PositionInterlock_APLC_Input[1].EquipmentInterlock_APLC_Input[1].SignalInterlock_APLC_Input[1] )
   END_RUNG
   RUNG wire#powerrail
      Contact( "Get Sinais de Interlock Falcare".Station[8]."Sinal do job"[1] )
      I_Contact( "BYPASS_MOD_1" )
      I_Contact( "BYPASS_GERAL" )
      I_Contact( "BYPASS_POSTO_60" )
      Coil( "Signals".ProcessInterlock_APLC_Input[1].ModezoneInterlock_APLC_Input[1].StationInterlock_APLC_Input[11].PositionInterlock_APLC_Input[1].EquipmentInterlock_APLC_Input[1].SignalInterlock_APLC_Input[2] )
   END_RUNG
   RUNG wire#powerrail
      I_Contact( "Get Sinais de Interlock Falcare".Station[8]."Sinal do job"[3] )
      I_Contact( "BYPASS_MOD_1" )
      I_Contact( "BYPASS_GERAL" )
      I_Contact( "BYPASS_POSTO_60" )
      Coil( "Signals".ProcessInterlock_APLC_Input[1].ModezoneInterlock_APLC_Input[1].StationInterlock_APLC_Input[11].PositionInterlock_APLC_Input[1].EquipmentInterlock_APLC_Input[2].SignalInterlock_APLC_Input[2] )
   END_RUNG
   RUNG wire#powerrail
      Contact( "Get Sinais de Interlock Falcare".Station[8]."Sinal do job"[4] )
      I_Contact( "BYPASS_MOD_1" )
      I_Contact( "BYPASS_GERAL" )
      I_Contact( "BYPASS_POSTO_60" )
      Coil( "Signals".ProcessInterlock_APLC_Input[1].ModezoneInterlock_APLC_Input[1].StationInterlock_APLC_Input[11].PositionInterlock_APLC_Input[1].EquipmentInterlock_APLC_Input[1].SignalInterlock_APLC_Input[3] )
   END_RUNG
   RUNG wire#powerrail
      Contact( "Get Sinais de Interlock Falcare".Station[8]."Sinal do job"[5] )
      I_Contact( "BYPASS_MOD_1" )
      I_Contact( "BYPASS_GERAL" )
      I_Contact( "Get Sinais de Interlock Falcare".Station[8]."Sinal do job"[6] )
      I_Contact( "BYPASS_POSTO_60" )
      Coil( "Signals".ProcessInterlock_APLC_Input[1].ModezoneInterlock_APLC_Input[1].StationInterlock_APLC_Input[11].PositionInterlock_APLC_Input[1].EquipmentInterlock_APLC_Input[1].SignalInterlock_APLC_Input[4] )
   END_RUNG
   RUNG wire#powerrail
      Contact( "Get Sinais de Interlock Falcare".Station[8]."Sinal do job"[6] )
      I_Contact( "BYPASS_MOD_1" )
      I_Contact( "BYPASS_GERAL" )
      I_Contact( "BYPASS_POSTO_60" )
      Coil( "Signals".ProcessInterlock_APLC_Input[1].ModezoneInterlock_APLC_Input[1].StationInterlock_APLC_Input[11].PositionInterlock_APLC_Input[1].EquipmentInterlock_APLC_Input[1].SignalInterlock_APLC_Input[5] )
   END_RUNG
   RUNG wire#powerrail
      Contact( "Get Sinais de Interlock Falcare".Station[8]."Sinal do job"[7] )
      I_Contact( "BYPASS_MOD_1" )
      I_Contact( "BYPASS_GERAL" )
      I_Contact( "BYPASS_POSTO_60" )
      Coil( "Signals".ProcessInterlock_APLC_Input[1].ModezoneInterlock_APLC_Input[1].StationInterlock_APLC_Input[11].PositionInterlock_APLC_Input[1].EquipmentInterlock_APLC_Input[1].SignalInterlock_APLC_Input[6] )
   END_RUNG
   RUNG wire#powerrail
      I_Contact( "Get Sinais de Interlock Falcare".Station[8]."Sinal do job"[9] )
      I_Contact( "BYPASS_MOD_1" )
      I_Contact( "BYPASS_GERAL" )
      I_Contact( "Put Sinais de Interlock Falcare".Bypass_Cortina )
      Coil( "Signals".ProcessInterlock_APLC_Input[1].ModezoneInterlock_APLC_Input[1].StationInterlock_APLC_Input[4].PositionInterlock_APLC_Input[1].EquipmentInterlock_APLC_Input[1].SignalInterlock_APLC_Input[6] )
   END_RUNG
   RUNG wire#powerrail
      I_Contact( "Get Sinais de Interlock Falcare".Station[8]."Sinal do job"[8] )
      I_Contact( "BYPASS_MOD_1" )
      I_Contact( "BYPASS_GERAL" )
      I_Contact( "Put Sinais de Interlock Falcare".Bypass_Cortina )
      Coil( "Signals".ProcessInterlock_APLC_Input[1].ModezoneInterlock_APLC_Input[1].StationInterlock_APLC_Input[4].PositionInterlock_APLC_Input[1].EquipmentInterlock_APLC_Input[1].SignalInterlock_APLC_Input[7] )
   END_RUNG
   RUNG wire#powerrail
      Contact( "AlwaysFALSE" )
      Coil( "Put Sinais de Interlock Falcare".Bypass_Cortina )
   END_RUNG
   // the same network as SCL:
   "Signals".ProcessInterlock_APLC_Input[1].ModezoneInterlock_APLC_Input[1].StationInterlock_APLC_Input[11].PositionInterlock_APLC_Input[1].EquipmentInterlock_APLC_Input[1].SignalInterlock_APLC_Input[1] := "Get Sinais de Interlock Falcare".Station[8]."Sinal do job"[0] AND NOT "BYPASS_MOD_1" AND NOT "BYPASS_GERAL" AND NOT "BYPASS_POSTO_60";
   "Signals".ProcessInterlock_APLC_Input[1].ModezoneInterlock_APLC_Input[1].StationInterlock_APLC_Input[11].PositionInterlock_APLC_Input[1].EquipmentInterlock_APLC_Input[1].SignalInterlock_APLC_Input[2] := "Get Sinais de Interlock Falcare".Station[8]."Sinal do job"[1] AND NOT "BYPASS_MOD_1" AND NOT "BYPASS_GERAL" AND NOT "BYPASS_POSTO_60";
   "Signals".ProcessInterlock_APLC_Input[1].ModezoneInterlock_APLC_Input[1].StationInterlock_APLC_Input[11].PositionInterlock_APLC_Input[1].EquipmentInterlock_APLC_Input[2].SignalInterlock_APLC_Input[2] := NOT "Get Sinais de Interlock Falcare".Station[8]."Sinal do job"[3] AND NOT "BYPASS_MOD_1" AND NOT "BYPASS_GERAL" AND NOT "BYPASS_POSTO_60";
   "Signals".ProcessInterlock_APLC_Input[1].ModezoneInterlock_APLC_Input[1].StationInterlock_APLC_Input[11].PositionInterlock_APLC_Input[1].EquipmentInterlock_APLC_Input[1].SignalInterlock_APLC_Input[3] := "Get Sinais de Interlock Falcare".Station[8]."Sinal do job"[4] AND NOT "BYPASS_MOD_1" AND NOT "BYPASS_GERAL" AND NOT "BYPASS_POSTO_60";
   "Signals".ProcessInterlock_APLC_Input[1].ModezoneInterlock_APLC_Input[1].StationInterlock_APLC_Input[11].PositionInterlock_APLC_Input[1].EquipmentInterlock_APLC_Input[1].SignalInterlock_APLC_Input[4] := "Get Sinais de Interlock Falcare".Station[8]."Sinal do job"[5] AND NOT "BYPASS_MOD_1" AND NOT "BYPASS_GERAL" AND NOT "Get Sinais de Interlock Falcare".Station[8]."Sinal do job"[6] AND NOT "BYPASS_POSTO_60";
   "Signals".ProcessInterlock_APLC_Input[1].ModezoneInterlock_APLC_Input[1].StationInterlock_APLC_Input[11].PositionInterlock_APLC_Input[1].EquipmentInterlock_APLC_Input[1].SignalInterlock_APLC_Input[5] := "Get Sinais de Interlock Falcare".Station[8]."Sinal do job"[6] AND NOT "BYPASS_MOD_1" AND NOT "BYPASS_GERAL" AND NOT "BYPASS_POSTO_60";
   "Signals".ProcessInterlock_APLC_Input[1].ModezoneInterlock_APLC_Input[1].StationInterlock_APLC_Input[11].PositionInterlock_APLC_Input[1].EquipmentInterlock_APLC_Input[1].SignalInterlock_APLC_Input[6] := "Get Sinais de Interlock Falcare".Station[8]."Sinal do job"[7] AND NOT "BYPASS_MOD_1" AND NOT "BYPASS_GERAL" AND NOT "BYPASS_POSTO_60";
   "Signals".ProcessInterlock_APLC_Input[1].ModezoneInterlock_APLC_Input[1].StationInterlock_APLC_Input[4].PositionInterlock_APLC_Input[1].EquipmentInterlock_APLC_Input[1].SignalInterlock_APLC_Input[6] := NOT "Get Sinais de Interlock Falcare".Station[8]."Sinal do job"[9] AND NOT "BYPASS_MOD_1" AND NOT "BYPASS_GERAL" AND NOT "Put Sinais de Interlock Falcare".Bypass_Cortina;
   "Signals".ProcessInterlock_APLC_Input[1].ModezoneInterlock_APLC_Input[1].StationInterlock_APLC_Input[4].PositionInterlock_APLC_Input[1].EquipmentInterlock_APLC_Input[1].SignalInterlock_APLC_Input[7] := NOT "Get Sinais de Interlock Falcare".Station[8]."Sinal do job"[8] AND NOT "BYPASS_MOD_1" AND NOT "BYPASS_GERAL" AND NOT "Put Sinais de Interlock Falcare".Bypass_Cortina;
   "Put Sinais de Interlock Falcare".Bypass_Cortina := "AlwaysFALSE";
END_REGION

REGION Network 13: ALARME IHM TRANSPORTADOR FALCARE
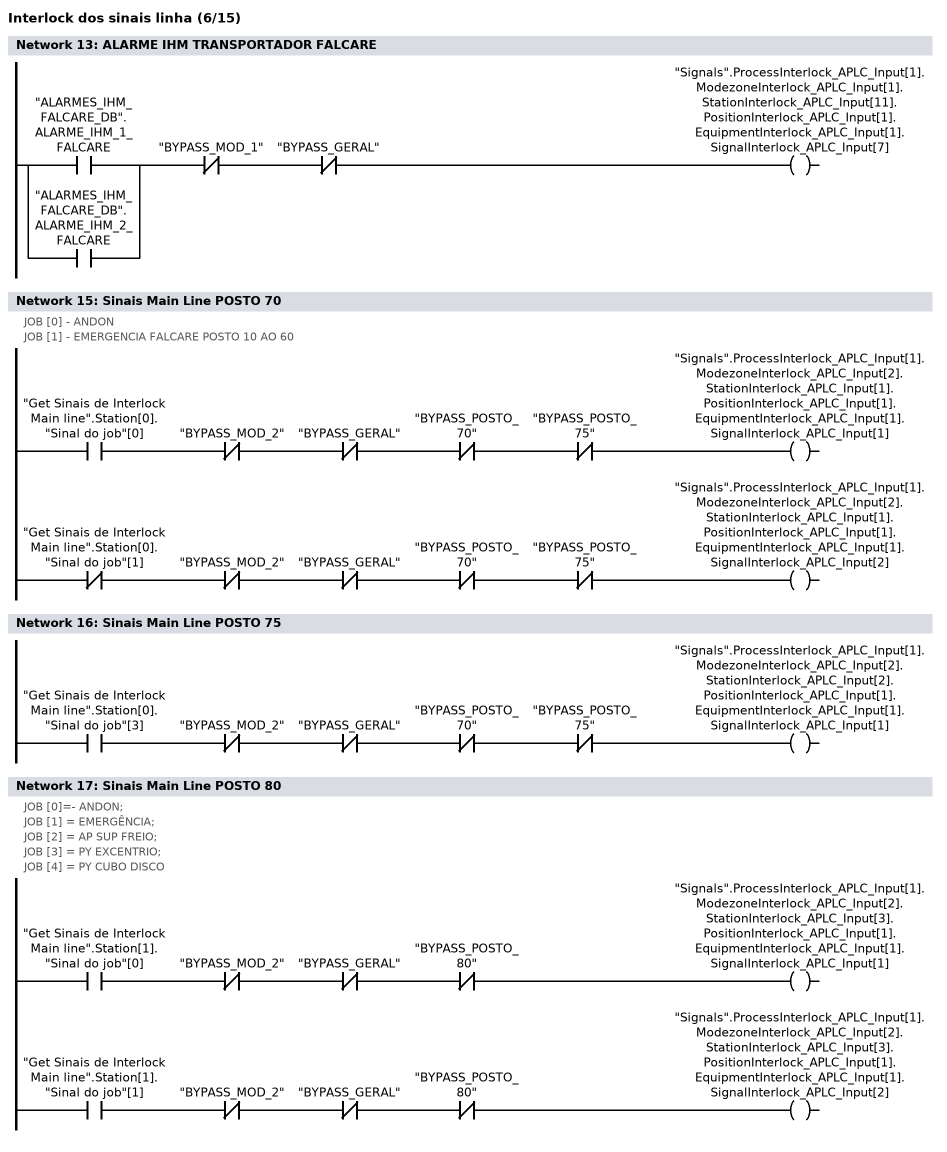
   RUNG wire#powerrail
      Contact( "ALARMES_IHM_FALCARE_DB".ALARME_IHM_1_FALCARE )
      wire#w1
      I_Contact( "BYPASS_MOD_1" )
      I_Contact( "BYPASS_GERAL" )
      Coil( "Signals".ProcessInterlock_APLC_Input[1].ModezoneInterlock_APLC_Input[1].StationInterlock_APLC_Input[11].PositionInterlock_APLC_Input[1].EquipmentInterlock_APLC_Input[1].SignalInterlock_APLC_Input[7] )
   END_RUNG
   RUNG wire#powerrail
      Contact( "ALARMES_IHM_FALCARE_DB".ALARME_IHM_2_FALCARE )
   END_RUNG wire#w1
   // the same network as SCL:
   "Signals".ProcessInterlock_APLC_Input[1].ModezoneInterlock_APLC_Input[1].StationInterlock_APLC_Input[11].PositionInterlock_APLC_Input[1].EquipmentInterlock_APLC_Input[1].SignalInterlock_APLC_Input[7] := ("ALARMES_IHM_FALCARE_DB".ALARME_IHM_1_FALCARE OR "ALARMES_IHM_FALCARE_DB".ALARME_IHM_2_FALCARE) AND NOT "BYPASS_MOD_1" AND NOT "BYPASS_GERAL";
END_REGION

REGION Network 14: Sinais GIRADOR
END_REGION

REGION Network 15: Sinais Main Line POSTO 70
   // JOB [0] - ANDON
   // JOB [1] - EMERGENCIA FALCARE POSTO 10 AO 60
   RUNG wire#powerrail
      Contact( "Get Sinais de Interlock Main line".Station[0]."Sinal do job"[0] )
      I_Contact( "BYPASS_MOD_2" )
      I_Contact( "BYPASS_GERAL" )
      I_Contact( "BYPASS_POSTO_70" )
      I_Contact( "BYPASS_POSTO_75" )
      Coil( "Signals".ProcessInterlock_APLC_Input[1].ModezoneInterlock_APLC_Input[2].StationInterlock_APLC_Input[1].PositionInterlock_APLC_Input[1].EquipmentInterlock_APLC_Input[1].SignalInterlock_APLC_Input[1] )
   END_RUNG
   RUNG wire#powerrail
      I_Contact( "Get Sinais de Interlock Main line".Station[0]."Sinal do job"[1] )
      I_Contact( "BYPASS_MOD_2" )
      I_Contact( "BYPASS_GERAL" )
      I_Contact( "BYPASS_POSTO_70" )
      I_Contact( "BYPASS_POSTO_75" )
      Coil( "Signals".ProcessInterlock_APLC_Input[1].ModezoneInterlock_APLC_Input[2].StationInterlock_APLC_Input[1].PositionInterlock_APLC_Input[1].EquipmentInterlock_APLC_Input[1].SignalInterlock_APLC_Input[2] )
   END_RUNG
   // the same network as SCL:
   "Signals".ProcessInterlock_APLC_Input[1].ModezoneInterlock_APLC_Input[2].StationInterlock_APLC_Input[1].PositionInterlock_APLC_Input[1].EquipmentInterlock_APLC_Input[1].SignalInterlock_APLC_Input[1] := "Get Sinais de Interlock Main line".Station[0]."Sinal do job"[0] AND NOT "BYPASS_MOD_2" AND NOT "BYPASS_GERAL" AND NOT "BYPASS_POSTO_70" AND NOT "BYPASS_POSTO_75";
   "Signals".ProcessInterlock_APLC_Input[1].ModezoneInterlock_APLC_Input[2].StationInterlock_APLC_Input[1].PositionInterlock_APLC_Input[1].EquipmentInterlock_APLC_Input[1].SignalInterlock_APLC_Input[2] := NOT "Get Sinais de Interlock Main line".Station[0]."Sinal do job"[1] AND NOT "BYPASS_MOD_2" AND NOT "BYPASS_GERAL" AND NOT "BYPASS_POSTO_70" AND NOT "BYPASS_POSTO_75";
END_REGION

REGION Network 16: Sinais Main Line POSTO 75
   RUNG wire#powerrail
      Contact( "Get Sinais de Interlock Main line".Station[0]."Sinal do job"[3] )
      I_Contact( "BYPASS_MOD_2" )
      I_Contact( "BYPASS_GERAL" )
      I_Contact( "BYPASS_POSTO_70" )
      I_Contact( "BYPASS_POSTO_75" )
      Coil( "Signals".ProcessInterlock_APLC_Input[1].ModezoneInterlock_APLC_Input[2].StationInterlock_APLC_Input[2].PositionInterlock_APLC_Input[1].EquipmentInterlock_APLC_Input[1].SignalInterlock_APLC_Input[1] )
   END_RUNG
   // the same network as SCL:
   "Signals".ProcessInterlock_APLC_Input[1].ModezoneInterlock_APLC_Input[2].StationInterlock_APLC_Input[2].PositionInterlock_APLC_Input[1].EquipmentInterlock_APLC_Input[1].SignalInterlock_APLC_Input[1] := "Get Sinais de Interlock Main line".Station[0]."Sinal do job"[3] AND NOT "BYPASS_MOD_2" AND NOT "BYPASS_GERAL" AND NOT "BYPASS_POSTO_70" AND NOT "BYPASS_POSTO_75";
END_REGION

REGION Network 17: Sinais Main Line POSTO 80
   // JOB [0]=- ANDON;
   // JOB [1] = EMERGÊNCIA;
   // JOB [2] = AP SUP FREIO;
   // JOB [3] = PY EXCENTRIO;
   // JOB [4] = PY CUBO DISCO
   RUNG wire#powerrail
      Contact( "Get Sinais de Interlock Main line".Station[1]."Sinal do job"[0] )
      I_Contact( "BYPASS_MOD_2" )
      I_Contact( "BYPASS_GERAL" )
      I_Contact( "BYPASS_POSTO_80" )
      Coil( "Signals".ProcessInterlock_APLC_Input[1].ModezoneInterlock_APLC_Input[2].StationInterlock_APLC_Input[3].PositionInterlock_APLC_Input[1].EquipmentInterlock_APLC_Input[1].SignalInterlock_APLC_Input[1] )
   END_RUNG
   RUNG wire#powerrail
      Contact( "Get Sinais de Interlock Main line".Station[1]."Sinal do job"[1] )
      I_Contact( "BYPASS_MOD_2" )
      I_Contact( "BYPASS_GERAL" )
      I_Contact( "BYPASS_POSTO_80" )
      Coil( "Signals".ProcessInterlock_APLC_Input[1].ModezoneInterlock_APLC_Input[2].StationInterlock_APLC_Input[3].PositionInterlock_APLC_Input[1].EquipmentInterlock_APLC_Input[1].SignalInterlock_APLC_Input[2] )
   END_RUNG
   // the same network as SCL:
   "Signals".ProcessInterlock_APLC_Input[1].ModezoneInterlock_APLC_Input[2].StationInterlock_APLC_Input[3].PositionInterlock_APLC_Input[1].EquipmentInterlock_APLC_Input[1].SignalInterlock_APLC_Input[1] := "Get Sinais de Interlock Main line".Station[1]."Sinal do job"[0] AND NOT "BYPASS_MOD_2" AND NOT "BYPASS_GERAL" AND NOT "BYPASS_POSTO_80";
   "Signals".ProcessInterlock_APLC_Input[1].ModezoneInterlock_APLC_Input[2].StationInterlock_APLC_Input[3].PositionInterlock_APLC_Input[1].EquipmentInterlock_APLC_Input[1].SignalInterlock_APLC_Input[2] := "Get Sinais de Interlock Main line".Station[1]."Sinal do job"[1] AND NOT "BYPASS_MOD_2" AND NOT "BYPASS_GERAL" AND NOT "BYPASS_POSTO_80";
END_REGION

REGION Network 18: Sinais Main Line POSTO 90
   // JOB [0] = ANDON;
   // JOB [1] = EMERGÊNCIA;
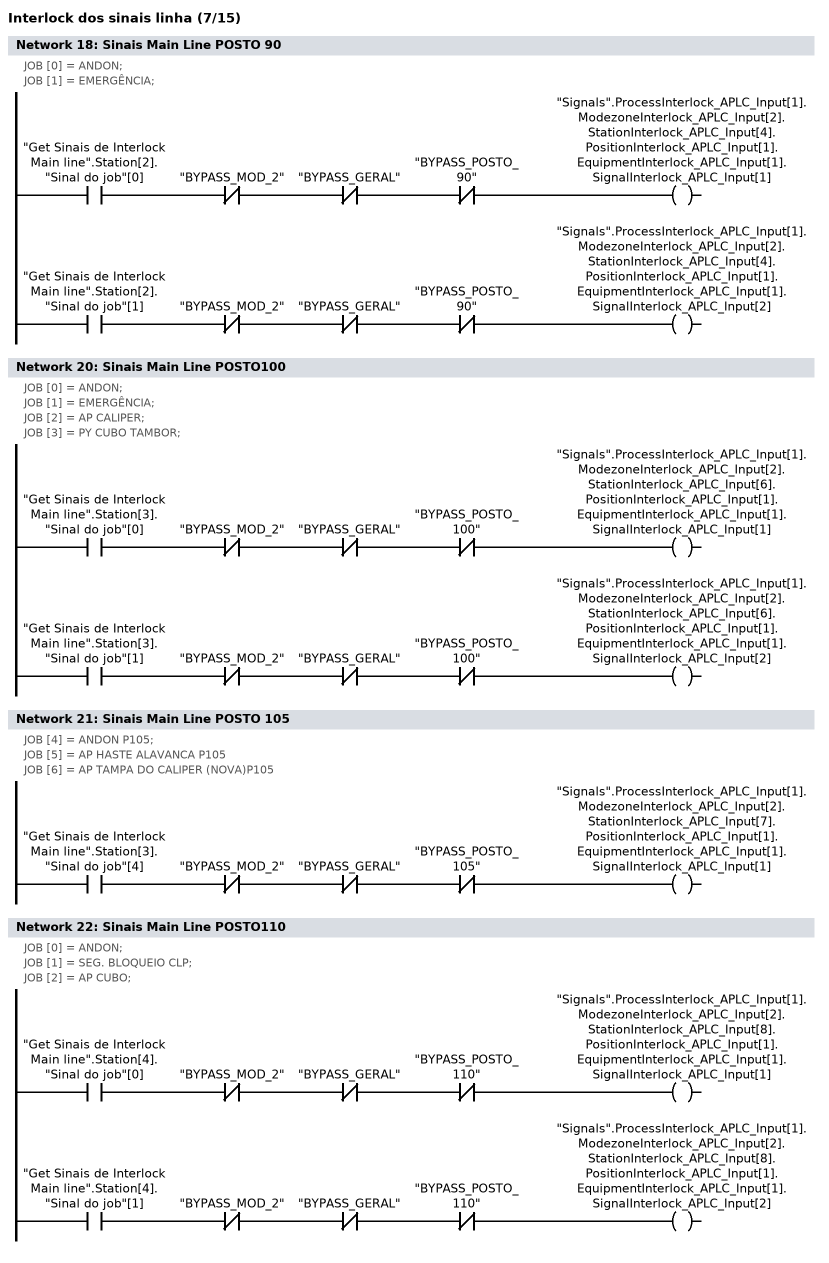
   RUNG wire#powerrail
      Contact( "Get Sinais de Interlock Main line".Station[2]."Sinal do job"[0] )
      I_Contact( "BYPASS_MOD_2" )
      I_Contact( "BYPASS_GERAL" )
      I_Contact( "BYPASS_POSTO_90" )
      Coil( "Signals".ProcessInterlock_APLC_Input[1].ModezoneInterlock_APLC_Input[2].StationInterlock_APLC_Input[4].PositionInterlock_APLC_Input[1].EquipmentInterlock_APLC_Input[1].SignalInterlock_APLC_Input[1] )
   END_RUNG
   RUNG wire#powerrail
      Contact( "Get Sinais de Interlock Main line".Station[2]."Sinal do job"[1] )
      I_Contact( "BYPASS_MOD_2" )
      I_Contact( "BYPASS_GERAL" )
      I_Contact( "BYPASS_POSTO_90" )
      Coil( "Signals".ProcessInterlock_APLC_Input[1].ModezoneInterlock_APLC_Input[2].StationInterlock_APLC_Input[4].PositionInterlock_APLC_Input[1].EquipmentInterlock_APLC_Input[1].SignalInterlock_APLC_Input[2] )
   END_RUNG
   // the same network as SCL:
   "Signals".ProcessInterlock_APLC_Input[1].ModezoneInterlock_APLC_Input[2].StationInterlock_APLC_Input[4].PositionInterlock_APLC_Input[1].EquipmentInterlock_APLC_Input[1].SignalInterlock_APLC_Input[1] := "Get Sinais de Interlock Main line".Station[2]."Sinal do job"[0] AND NOT "BYPASS_MOD_2" AND NOT "BYPASS_GERAL" AND NOT "BYPASS_POSTO_90";
   "Signals".ProcessInterlock_APLC_Input[1].ModezoneInterlock_APLC_Input[2].StationInterlock_APLC_Input[4].PositionInterlock_APLC_Input[1].EquipmentInterlock_APLC_Input[1].SignalInterlock_APLC_Input[2] := "Get Sinais de Interlock Main line".Station[2]."Sinal do job"[1] AND NOT "BYPASS_MOD_2" AND NOT "BYPASS_GERAL" AND NOT "BYPASS_POSTO_90";
END_REGION

REGION Network 19: Sinais Main Line POSTO 95
   // JOB [2] = AP HOLDER. P95
END_REGION

REGION Network 20: Sinais Main Line POSTO100
   // JOB [0] = ANDON;
   // JOB [1] = EMERGÊNCIA;
   // JOB [2] = AP CALIPER;
   // JOB [3] = PY CUBO TAMBOR;
   RUNG wire#powerrail
      Contact( "Get Sinais de Interlock Main line".Station[3]."Sinal do job"[0] )
      I_Contact( "BYPASS_MOD_2" )
      I_Contact( "BYPASS_GERAL" )
      I_Contact( "BYPASS_POSTO_100" )
      Coil( "Signals".ProcessInterlock_APLC_Input[1].ModezoneInterlock_APLC_Input[2].StationInterlock_APLC_Input[6].PositionInterlock_APLC_Input[1].EquipmentInterlock_APLC_Input[1].SignalInterlock_APLC_Input[1] )
   END_RUNG
   RUNG wire#powerrail
      Contact( "Get Sinais de Interlock Main line".Station[3]."Sinal do job"[1] )
      I_Contact( "BYPASS_MOD_2" )
      I_Contact( "BYPASS_GERAL" )
      I_Contact( "BYPASS_POSTO_100" )
      Coil( "Signals".ProcessInterlock_APLC_Input[1].ModezoneInterlock_APLC_Input[2].StationInterlock_APLC_Input[6].PositionInterlock_APLC_Input[1].EquipmentInterlock_APLC_Input[1].SignalInterlock_APLC_Input[2] )
   END_RUNG
   // the same network as SCL:
   "Signals".ProcessInterlock_APLC_Input[1].ModezoneInterlock_APLC_Input[2].StationInterlock_APLC_Input[6].PositionInterlock_APLC_Input[1].EquipmentInterlock_APLC_Input[1].SignalInterlock_APLC_Input[1] := "Get Sinais de Interlock Main line".Station[3]."Sinal do job"[0] AND NOT "BYPASS_MOD_2" AND NOT "BYPASS_GERAL" AND NOT "BYPASS_POSTO_100";
   "Signals".ProcessInterlock_APLC_Input[1].ModezoneInterlock_APLC_Input[2].StationInterlock_APLC_Input[6].PositionInterlock_APLC_Input[1].EquipmentInterlock_APLC_Input[1].SignalInterlock_APLC_Input[2] := "Get Sinais de Interlock Main line".Station[3]."Sinal do job"[1] AND NOT "BYPASS_MOD_2" AND NOT "BYPASS_GERAL" AND NOT "BYPASS_POSTO_100";
END_REGION

REGION Network 21: Sinais Main Line POSTO 105
   // JOB [4] = ANDON P105;
   // JOB [5] = AP HASTE ALAVANCA P105
   // JOB [6] = AP TAMPA DO CALIPER (NOVA)P105
   RUNG wire#powerrail
      Contact( "Get Sinais de Interlock Main line".Station[3]."Sinal do job"[4] )
      I_Contact( "BYPASS_MOD_2" )
      I_Contact( "BYPASS_GERAL" )
      I_Contact( "BYPASS_POSTO_105" )
      Coil( "Signals".ProcessInterlock_APLC_Input[1].ModezoneInterlock_APLC_Input[2].StationInterlock_APLC_Input[7].PositionInterlock_APLC_Input[1].EquipmentInterlock_APLC_Input[1].SignalInterlock_APLC_Input[1] )
   END_RUNG
   // the same network as SCL:
   "Signals".ProcessInterlock_APLC_Input[1].ModezoneInterlock_APLC_Input[2].StationInterlock_APLC_Input[7].PositionInterlock_APLC_Input[1].EquipmentInterlock_APLC_Input[1].SignalInterlock_APLC_Input[1] := "Get Sinais de Interlock Main line".Station[3]."Sinal do job"[4] AND NOT "BYPASS_MOD_2" AND NOT "BYPASS_GERAL" AND NOT "BYPASS_POSTO_105";
END_REGION

REGION Network 22: Sinais Main Line POSTO110
   // JOB [0] = ANDON;
   // JOB [1] = SEG. BLOQUEIO CLP;
   // JOB [2] = AP CUBO;
   RUNG wire#powerrail
      Contact( "Get Sinais de Interlock Main line".Station[4]."Sinal do job"[0] )
      I_Contact( "BYPASS_MOD_2" )
      I_Contact( "BYPASS_GERAL" )
      I_Contact( "BYPASS_POSTO_110" )
      Coil( "Signals".ProcessInterlock_APLC_Input[1].ModezoneInterlock_APLC_Input[2].StationInterlock_APLC_Input[8].PositionInterlock_APLC_Input[1].EquipmentInterlock_APLC_Input[1].SignalInterlock_APLC_Input[1] )
   END_RUNG
   RUNG wire#powerrail
      Contact( "Get Sinais de Interlock Main line".Station[4]."Sinal do job"[1] )
      I_Contact( "BYPASS_MOD_2" )
      I_Contact( "BYPASS_GERAL" )
      I_Contact( "BYPASS_POSTO_110" )
      Coil( "Signals".ProcessInterlock_APLC_Input[1].ModezoneInterlock_APLC_Input[2].StationInterlock_APLC_Input[8].PositionInterlock_APLC_Input[1].EquipmentInterlock_APLC_Input[1].SignalInterlock_APLC_Input[2] )
   END_RUNG
   // the same network as SCL:
   "Signals".ProcessInterlock_APLC_Input[1].ModezoneInterlock_APLC_Input[2].StationInterlock_APLC_Input[8].PositionInterlock_APLC_Input[1].EquipmentInterlock_APLC_Input[1].SignalInterlock_APLC_Input[1] := "Get Sinais de Interlock Main line".Station[4]."Sinal do job"[0] AND NOT "BYPASS_MOD_2" AND NOT "BYPASS_GERAL" AND NOT "BYPASS_POSTO_110";
   "Signals".ProcessInterlock_APLC_Input[1].ModezoneInterlock_APLC_Input[2].StationInterlock_APLC_Input[8].PositionInterlock_APLC_Input[1].EquipmentInterlock_APLC_Input[1].SignalInterlock_APLC_Input[2] := "Get Sinais de Interlock Main line".Station[4]."Sinal do job"[1] AND NOT "BYPASS_MOD_2" AND NOT "BYPASS_GERAL" AND NOT "BYPASS_POSTO_110";
END_REGION

REGION Network 23: Sinais Main Line POSTO 115
   // JOB [3] = ANDON P115;
   // JOB [4] = CRAVADOR.
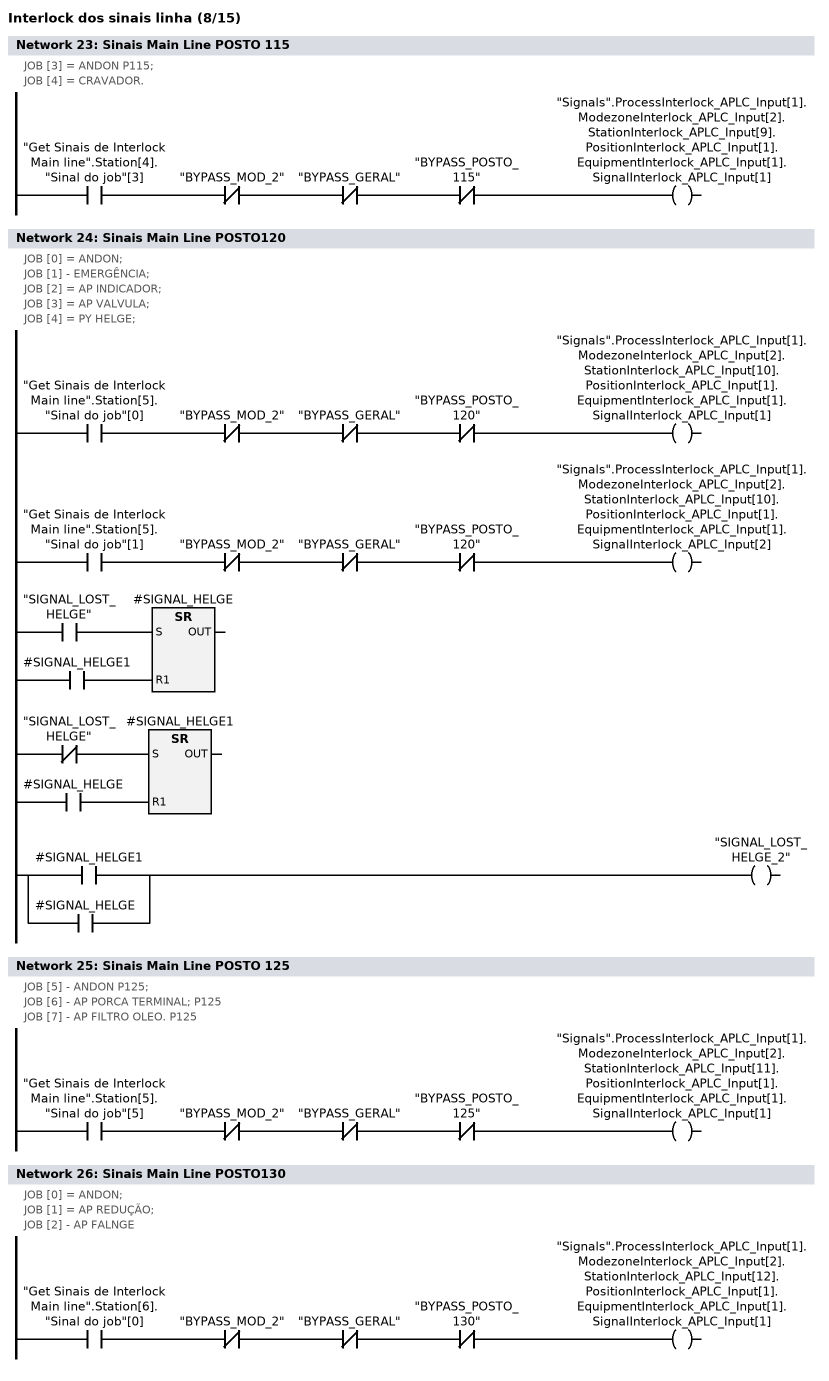
   RUNG wire#powerrail
      Contact( "Get Sinais de Interlock Main line".Station[4]."Sinal do job"[3] )
      I_Contact( "BYPASS_MOD_2" )
      I_Contact( "BYPASS_GERAL" )
      I_Contact( "BYPASS_POSTO_115" )
      Coil( "Signals".ProcessInterlock_APLC_Input[1].ModezoneInterlock_APLC_Input[2].StationInterlock_APLC_Input[9].PositionInterlock_APLC_Input[1].EquipmentInterlock_APLC_Input[1].SignalInterlock_APLC_Input[1] )
   END_RUNG
   // the same network as SCL:
   "Signals".ProcessInterlock_APLC_Input[1].ModezoneInterlock_APLC_Input[2].StationInterlock_APLC_Input[9].PositionInterlock_APLC_Input[1].EquipmentInterlock_APLC_Input[1].SignalInterlock_APLC_Input[1] := "Get Sinais de Interlock Main line".Station[4]."Sinal do job"[3] AND NOT "BYPASS_MOD_2" AND NOT "BYPASS_GERAL" AND NOT "BYPASS_POSTO_115";
END_REGION

REGION Network 24: Sinais Main Line POSTO120
   // JOB [0] = ANDON;
   // JOB [1] - EMERGÊNCIA;
   // JOB [2] = AP INDICADOR;
   // JOB [3] = AP VALVULA;
   // JOB [4] = PY HELGE;
   RUNG wire#powerrail
      Contact( "Get Sinais de Interlock Main line".Station[5]."Sinal do job"[0] )
      I_Contact( "BYPASS_MOD_2" )
      I_Contact( "BYPASS_GERAL" )
      I_Contact( "BYPASS_POSTO_120" )
      Coil( "Signals".ProcessInterlock_APLC_Input[1].ModezoneInterlock_APLC_Input[2].StationInterlock_APLC_Input[10].PositionInterlock_APLC_Input[1].EquipmentInterlock_APLC_Input[1].SignalInterlock_APLC_Input[1] )
   END_RUNG
   RUNG wire#powerrail
      Contact( "Get Sinais de Interlock Main line".Station[5]."Sinal do job"[1] )
      I_Contact( "BYPASS_MOD_2" )
      I_Contact( "BYPASS_GERAL" )
      I_Contact( "BYPASS_POSTO_120" )
      Coil( "Signals".ProcessInterlock_APLC_Input[1].ModezoneInterlock_APLC_Input[2].StationInterlock_APLC_Input[10].PositionInterlock_APLC_Input[1].EquipmentInterlock_APLC_Input[1].SignalInterlock_APLC_Input[2] )
   END_RUNG
   RUNG wire#powerrail
      Contact( "SIGNAL_LOST_HELGE" )
      S_SR(operand := #SIGNAL_HELGE, r1 := wire#w1)
   END_RUNG
   RUNG wire#powerrail
      Contact( #SIGNAL_HELGE1 )
   END_RUNG wire#w1
   RUNG wire#powerrail
      I_Contact( "SIGNAL_LOST_HELGE" )
      S_SR(operand := #SIGNAL_HELGE1, r1 := wire#w2)
   END_RUNG
   RUNG wire#powerrail
      Contact( #SIGNAL_HELGE )
   END_RUNG wire#w2
   RUNG wire#powerrail
      Contact( #SIGNAL_HELGE1 )
      wire#w3
      Coil( "SIGNAL_LOST_HELGE_2" )
   END_RUNG
   RUNG wire#powerrail
      Contact( #SIGNAL_HELGE )
   END_RUNG wire#w3
   // the same network as SCL:
   "Signals".ProcessInterlock_APLC_Input[1].ModezoneInterlock_APLC_Input[2].StationInterlock_APLC_Input[10].PositionInterlock_APLC_Input[1].EquipmentInterlock_APLC_Input[1].SignalInterlock_APLC_Input[1] := "Get Sinais de Interlock Main line".Station[5]."Sinal do job"[0] AND NOT "BYPASS_MOD_2" AND NOT "BYPASS_GERAL" AND NOT "BYPASS_POSTO_120";
   "Signals".ProcessInterlock_APLC_Input[1].ModezoneInterlock_APLC_Input[2].StationInterlock_APLC_Input[10].PositionInterlock_APLC_Input[1].EquipmentInterlock_APLC_Input[1].SignalInterlock_APLC_Input[2] := "Get Sinais de Interlock Main line".Station[5]."Sinal do job"[1] AND NOT "BYPASS_MOD_2" AND NOT "BYPASS_GERAL" AND NOT "BYPASS_POSTO_120";
   IF "SIGNAL_LOST_HELGE" THEN
       #SIGNAL_HELGE := TRUE;   // SR flip-flop
   END_IF;
   IF #SIGNAL_HELGE1 THEN #SIGNAL_HELGE := FALSE; END_IF;
   IF NOT "SIGNAL_LOST_HELGE" THEN
       #SIGNAL_HELGE1 := TRUE;   // SR flip-flop
   END_IF;
   IF #SIGNAL_HELGE THEN #SIGNAL_HELGE1 := FALSE; END_IF;
   "SIGNAL_LOST_HELGE_2" := #SIGNAL_HELGE1 OR #SIGNAL_HELGE;
END_REGION

REGION Network 25: Sinais Main Line POSTO 125
   // JOB [5] - ANDON P125;
   // JOB [6] - AP PORCA TERMINAL; P125
   // JOB [7] - AP FILTRO OLEO. P125
   RUNG wire#powerrail
      Contact( "Get Sinais de Interlock Main line".Station[5]."Sinal do job"[5] )
      I_Contact( "BYPASS_MOD_2" )
      I_Contact( "BYPASS_GERAL" )
      I_Contact( "BYPASS_POSTO_125" )
      Coil( "Signals".ProcessInterlock_APLC_Input[1].ModezoneInterlock_APLC_Input[2].StationInterlock_APLC_Input[11].PositionInterlock_APLC_Input[1].EquipmentInterlock_APLC_Input[1].SignalInterlock_APLC_Input[1] )
   END_RUNG
   // the same network as SCL:
   "Signals".ProcessInterlock_APLC_Input[1].ModezoneInterlock_APLC_Input[2].StationInterlock_APLC_Input[11].PositionInterlock_APLC_Input[1].EquipmentInterlock_APLC_Input[1].SignalInterlock_APLC_Input[1] := "Get Sinais de Interlock Main line".Station[5]."Sinal do job"[5] AND NOT "BYPASS_MOD_2" AND NOT "BYPASS_GERAL" AND NOT "BYPASS_POSTO_125";
END_REGION

REGION Network 26: Sinais Main Line POSTO130
   // JOB [0] = ANDON;
   // JOB [1] = AP REDUÇÃO;
   // JOB [2] - AP FALNGE
   RUNG wire#powerrail
      Contact( "Get Sinais de Interlock Main line".Station[6]."Sinal do job"[0] )
      I_Contact( "BYPASS_MOD_2" )
      I_Contact( "BYPASS_GERAL" )
      I_Contact( "BYPASS_POSTO_130" )
      Coil( "Signals".ProcessInterlock_APLC_Input[1].ModezoneInterlock_APLC_Input[2].StationInterlock_APLC_Input[12].PositionInterlock_APLC_Input[1].EquipmentInterlock_APLC_Input[1].SignalInterlock_APLC_Input[1] )
   END_RUNG
   // the same network as SCL:
   "Signals".ProcessInterlock_APLC_Input[1].ModezoneInterlock_APLC_Input[2].StationInterlock_APLC_Input[12].PositionInterlock_APLC_Input[1].EquipmentInterlock_APLC_Input[1].SignalInterlock_APLC_Input[1] := "Get Sinais de Interlock Main line".Station[6]."Sinal do job"[0] AND NOT "BYPASS_MOD_2" AND NOT "BYPASS_GERAL" AND NOT "BYPASS_POSTO_130";
END_REGION

REGION Network 27: Sinais Main Line POSTO140
   // JOB [0] = ANDON;
   // JOB [1] = EMERGÊNCIA;
   // JOB [2] = ESTANQUEIDADE CILINDRO;
   // JOB [3] = ESTANQUEIDADE CARCAÇA.
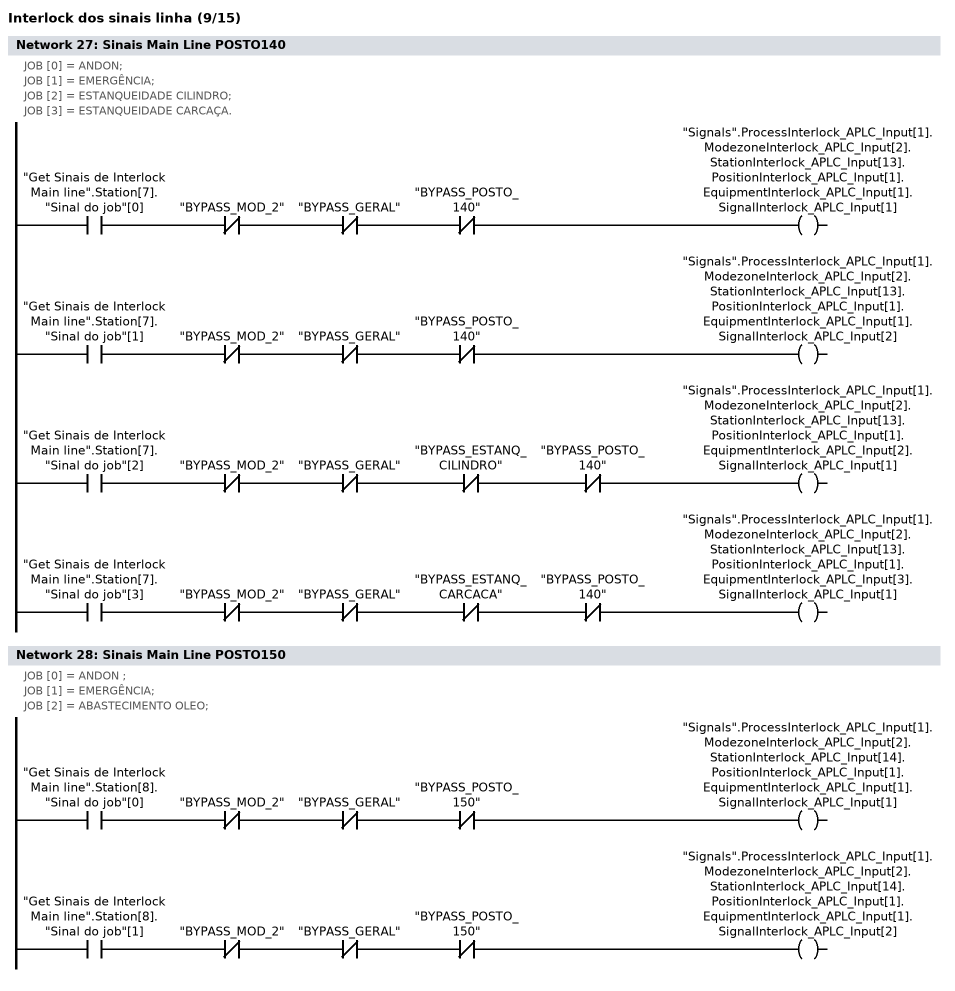
   RUNG wire#powerrail
      Contact( "Get Sinais de Interlock Main line".Station[7]."Sinal do job"[0] )
      I_Contact( "BYPASS_MOD_2" )
      I_Contact( "BYPASS_GERAL" )
      I_Contact( "BYPASS_POSTO_140" )
      Coil( "Signals".ProcessInterlock_APLC_Input[1].ModezoneInterlock_APLC_Input[2].StationInterlock_APLC_Input[13].PositionInterlock_APLC_Input[1].EquipmentInterlock_APLC_Input[1].SignalInterlock_APLC_Input[1] )
   END_RUNG
   RUNG wire#powerrail
      Contact( "Get Sinais de Interlock Main line".Station[7]."Sinal do job"[1] )
      I_Contact( "BYPASS_MOD_2" )
      I_Contact( "BYPASS_GERAL" )
      I_Contact( "BYPASS_POSTO_140" )
      Coil( "Signals".ProcessInterlock_APLC_Input[1].ModezoneInterlock_APLC_Input[2].StationInterlock_APLC_Input[13].PositionInterlock_APLC_Input[1].EquipmentInterlock_APLC_Input[1].SignalInterlock_APLC_Input[2] )
   END_RUNG
   RUNG wire#powerrail
      Contact( "Get Sinais de Interlock Main line".Station[7]."Sinal do job"[2] )
      I_Contact( "BYPASS_MOD_2" )
      I_Contact( "BYPASS_GERAL" )
      I_Contact( "BYPASS_ESTANQ_CILINDRO" )
      I_Contact( "BYPASS_POSTO_140" )
      Coil( "Signals".ProcessInterlock_APLC_Input[1].ModezoneInterlock_APLC_Input[2].StationInterlock_APLC_Input[13].PositionInterlock_APLC_Input[1].EquipmentInterlock_APLC_Input[2].SignalInterlock_APLC_Input[1] )
   END_RUNG
   RUNG wire#powerrail
      Contact( "Get Sinais de Interlock Main line".Station[7]."Sinal do job"[3] )
      I_Contact( "BYPASS_MOD_2" )
      I_Contact( "BYPASS_GERAL" )
      I_Contact( "BYPASS_ESTANQ_CARCACA" )
      I_Contact( "BYPASS_POSTO_140" )
      Coil( "Signals".ProcessInterlock_APLC_Input[1].ModezoneInterlock_APLC_Input[2].StationInterlock_APLC_Input[13].PositionInterlock_APLC_Input[1].EquipmentInterlock_APLC_Input[3].SignalInterlock_APLC_Input[1] )
   END_RUNG
   // the same network as SCL:
   "Signals".ProcessInterlock_APLC_Input[1].ModezoneInterlock_APLC_Input[2].StationInterlock_APLC_Input[13].PositionInterlock_APLC_Input[1].EquipmentInterlock_APLC_Input[1].SignalInterlock_APLC_Input[1] := "Get Sinais de Interlock Main line".Station[7]."Sinal do job"[0] AND NOT "BYPASS_MOD_2" AND NOT "BYPASS_GERAL" AND NOT "BYPASS_POSTO_140";
   "Signals".ProcessInterlock_APLC_Input[1].ModezoneInterlock_APLC_Input[2].StationInterlock_APLC_Input[13].PositionInterlock_APLC_Input[1].EquipmentInterlock_APLC_Input[1].SignalInterlock_APLC_Input[2] := "Get Sinais de Interlock Main line".Station[7]."Sinal do job"[1] AND NOT "BYPASS_MOD_2" AND NOT "BYPASS_GERAL" AND NOT "BYPASS_POSTO_140";
   "Signals".ProcessInterlock_APLC_Input[1].ModezoneInterlock_APLC_Input[2].StationInterlock_APLC_Input[13].PositionInterlock_APLC_Input[1].EquipmentInterlock_APLC_Input[2].SignalInterlock_APLC_Input[1] := "Get Sinais de Interlock Main line".Station[7]."Sinal do job"[2] AND NOT "BYPASS_MOD_2" AND NOT "BYPASS_GERAL" AND NOT "BYPASS_ESTANQ_CILINDRO" AND NOT "BYPASS_POSTO_140";
   "Signals".ProcessInterlock_APLC_Input[1].ModezoneInterlock_APLC_Input[2].StationInterlock_APLC_Input[13].PositionInterlock_APLC_Input[1].EquipmentInterlock_APLC_Input[3].SignalInterlock_APLC_Input[1] := "Get Sinais de Interlock Main line".Station[7]."Sinal do job"[3] AND NOT "BYPASS_MOD_2" AND NOT "BYPASS_GERAL" AND NOT "BYPASS_ESTANQ_CARCACA" AND NOT "BYPASS_POSTO_140";
END_REGION

REGION Network 28: Sinais Main Line POSTO150
   // JOB [0] = ANDON ;
   // JOB [1] = EMERGÊNCIA;
   // JOB [2] = ABASTECIMENTO OLEO;
   RUNG wire#powerrail
      Contact( "Get Sinais de Interlock Main line".Station[8]."Sinal do job"[0] )
      I_Contact( "BYPASS_MOD_2" )
      I_Contact( "BYPASS_GERAL" )
      I_Contact( "BYPASS_POSTO_150" )
      Coil( "Signals".ProcessInterlock_APLC_Input[1].ModezoneInterlock_APLC_Input[2].StationInterlock_APLC_Input[14].PositionInterlock_APLC_Input[1].EquipmentInterlock_APLC_Input[1].SignalInterlock_APLC_Input[1] )
   END_RUNG
   RUNG wire#powerrail
      Contact( "Get Sinais de Interlock Main line".Station[8]."Sinal do job"[1] )
      I_Contact( "BYPASS_MOD_2" )
      I_Contact( "BYPASS_GERAL" )
      I_Contact( "BYPASS_POSTO_150" )
      Coil( "Signals".ProcessInterlock_APLC_Input[1].ModezoneInterlock_APLC_Input[2].StationInterlock_APLC_Input[14].PositionInterlock_APLC_Input[1].EquipmentInterlock_APLC_Input[1].SignalInterlock_APLC_Input[2] )
   END_RUNG
   // the same network as SCL:
   "Signals".ProcessInterlock_APLC_Input[1].ModezoneInterlock_APLC_Input[2].StationInterlock_APLC_Input[14].PositionInterlock_APLC_Input[1].EquipmentInterlock_APLC_Input[1].SignalInterlock_APLC_Input[1] := "Get Sinais de Interlock Main line".Station[8]."Sinal do job"[0] AND NOT "BYPASS_MOD_2" AND NOT "BYPASS_GERAL" AND NOT "BYPASS_POSTO_150";
   "Signals".ProcessInterlock_APLC_Input[1].ModezoneInterlock_APLC_Input[2].StationInterlock_APLC_Input[14].PositionInterlock_APLC_Input[1].EquipmentInterlock_APLC_Input[1].SignalInterlock_APLC_Input[2] := "Get Sinais de Interlock Main line".Station[8]."Sinal do job"[1] AND NOT "BYPASS_MOD_2" AND NOT "BYPASS_GERAL" AND NOT "BYPASS_POSTO_150";
END_REGION

REGION Network 29: Sinais Main Line Q.G
   // JOB [0] = ANDON;
   // JOB [1] = EMERGÊNCIA;
   // JOB [2] - EIXO PENDURADO;
   // JOB [3] - GAP PRESENTE CAB;
   // JOB [4] - GAP PRESENTE TAKT 
   // STATION 10 JOB [0] = TRANSPORTADOR EM MANUAL
   // GAP + EIXO PENDURADO
   // MODEZONE 1 PARADO (FALCARE)
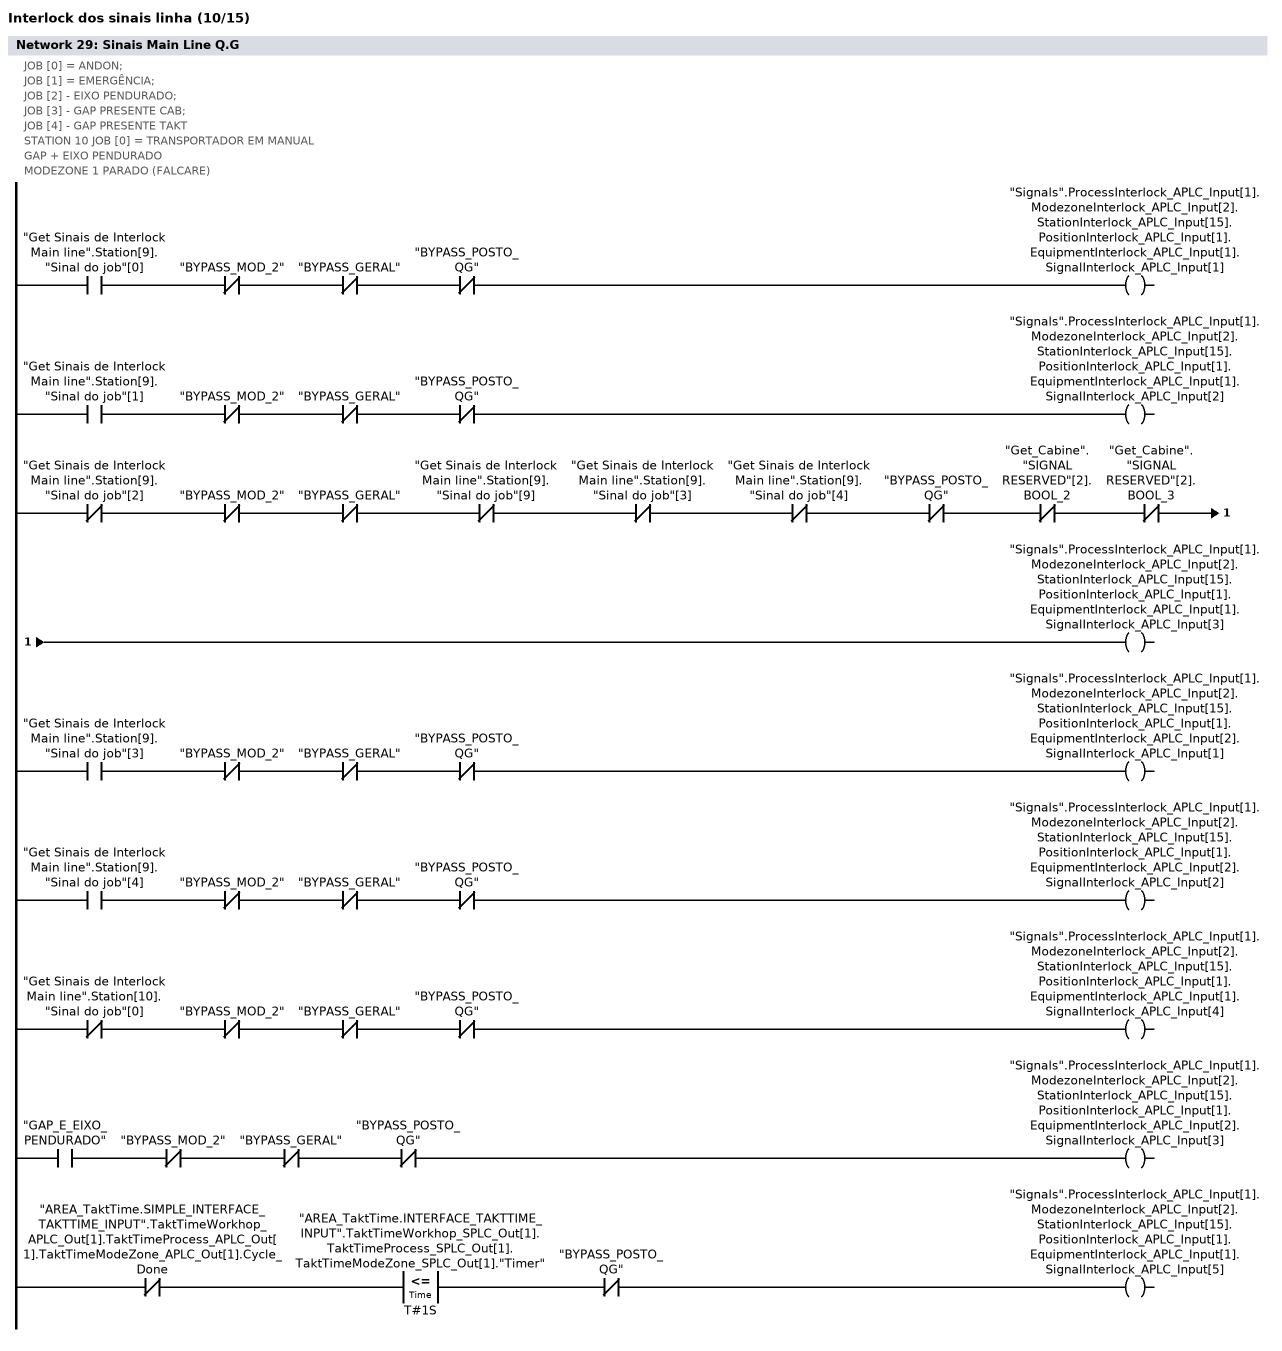
   RUNG wire#powerrail
      Contact( "Get Sinais de Interlock Main line".Station[9]."Sinal do job"[0] )
      I_Contact( "BYPASS_MOD_2" )
      I_Contact( "BYPASS_GERAL" )
      I_Contact( "BYPASS_POSTO_QG" )
      Coil( "Signals".ProcessInterlock_APLC_Input[1].ModezoneInterlock_APLC_Input[2].StationInterlock_APLC_Input[15].PositionInterlock_APLC_Input[1].EquipmentInterlock_APLC_Input[1].SignalInterlock_APLC_Input[1] )
   END_RUNG
   RUNG wire#powerrail
      Contact( "Get Sinais de Interlock Main line".Station[9]."Sinal do job"[1] )
      I_Contact( "BYPASS_MOD_2" )
      I_Contact( "BYPASS_GERAL" )
      I_Contact( "BYPASS_POSTO_QG" )
      Coil( "Signals".ProcessInterlock_APLC_Input[1].ModezoneInterlock_APLC_Input[2].StationInterlock_APLC_Input[15].PositionInterlock_APLC_Input[1].EquipmentInterlock_APLC_Input[1].SignalInterlock_APLC_Input[2] )
   END_RUNG
   RUNG wire#powerrail
      I_Contact( "Get Sinais de Interlock Main line".Station[9]."Sinal do job"[2] )
      I_Contact( "BYPASS_MOD_2" )
      I_Contact( "BYPASS_GERAL" )
      I_Contact( "Get Sinais de Interlock Main line".Station[9]."Sinal do job"[9] )
      I_Contact( "Get Sinais de Interlock Main line".Station[9]."Sinal do job"[3] )
      I_Contact( "Get Sinais de Interlock Main line".Station[9]."Sinal do job"[4] )
      I_Contact( "BYPASS_POSTO_QG" )
      I_Contact( "Get_Cabine"."SIGNAL RESERVED"[2].BOOL_2 )
      I_Contact( "Get_Cabine"."SIGNAL RESERVED"[2].BOOL_3 )
      Coil( "Signals".ProcessInterlock_APLC_Input[1].ModezoneInterlock_APLC_Input[2].StationInterlock_APLC_Input[15].PositionInterlock_APLC_Input[1].EquipmentInterlock_APLC_Input[1].SignalInterlock_APLC_Input[3] )
   END_RUNG
   RUNG wire#powerrail
      Contact( "Get Sinais de Interlock Main line".Station[9]."Sinal do job"[3] )
      I_Contact( "BYPASS_MOD_2" )
      I_Contact( "BYPASS_GERAL" )
      I_Contact( "BYPASS_POSTO_QG" )
      Coil( "Signals".ProcessInterlock_APLC_Input[1].ModezoneInterlock_APLC_Input[2].StationInterlock_APLC_Input[15].PositionInterlock_APLC_Input[1].EquipmentInterlock_APLC_Input[2].SignalInterlock_APLC_Input[1] )
   END_RUNG
   RUNG wire#powerrail
      Contact( "Get Sinais de Interlock Main line".Station[9]."Sinal do job"[4] )
      I_Contact( "BYPASS_MOD_2" )
      I_Contact( "BYPASS_GERAL" )
      I_Contact( "BYPASS_POSTO_QG" )
      Coil( "Signals".ProcessInterlock_APLC_Input[1].ModezoneInterlock_APLC_Input[2].StationInterlock_APLC_Input[15].PositionInterlock_APLC_Input[1].EquipmentInterlock_APLC_Input[2].SignalInterlock_APLC_Input[2] )
   END_RUNG
   RUNG wire#powerrail
      I_Contact( "Get Sinais de Interlock Main line".Station[10]."Sinal do job"[0] )
      I_Contact( "BYPASS_MOD_2" )
      I_Contact( "BYPASS_GERAL" )
      I_Contact( "BYPASS_POSTO_QG" )
      Coil( "Signals".ProcessInterlock_APLC_Input[1].ModezoneInterlock_APLC_Input[2].StationInterlock_APLC_Input[15].PositionInterlock_APLC_Input[1].EquipmentInterlock_APLC_Input[1].SignalInterlock_APLC_Input[4] )
   END_RUNG
   RUNG wire#powerrail
      Contact( "GAP_E_EIXO_PENDURADO" )
      I_Contact( "BYPASS_MOD_2" )
      I_Contact( "BYPASS_GERAL" )
      I_Contact( "BYPASS_POSTO_QG" )
      Coil( "Signals".ProcessInterlock_APLC_Input[1].ModezoneInterlock_APLC_Input[2].StationInterlock_APLC_Input[15].PositionInterlock_APLC_Input[1].EquipmentInterlock_APLC_Input[2].SignalInterlock_APLC_Input[3] )
   END_RUNG
   RUNG wire#powerrail
      I_Contact( "AREA_TaktTime.SIMPLE_INTERFACE_TAKTTIME_INPUT".TaktTimeWorkhop_APLC_Out[1].TaktTimeProcess_APLC_Out[1].TaktTimeModeZone_APLC_Out[1].Cycle_Done )
      { S7_Templates := "SrcType := Time" } LE_Contact(in1 := "AREA_TaktTime.INTERFACE_TAKTTIME_INPUT".TaktTimeWorkhop_SPLC_Out[1].TaktTimeProcess_SPLC_Out[1].TaktTimeModeZone_SPLC_Out[1]."Timer", in2 := T#1S)
      I_Contact( "BYPASS_POSTO_QG" )
      Coil( "Signals".ProcessInterlock_APLC_Input[1].ModezoneInterlock_APLC_Input[2].StationInterlock_APLC_Input[15].PositionInterlock_APLC_Input[1].EquipmentInterlock_APLC_Input[1].SignalInterlock_APLC_Input[5] )
   END_RUNG
   // the same network as SCL:
   "Signals".ProcessInterlock_APLC_Input[1].ModezoneInterlock_APLC_Input[2].StationInterlock_APLC_Input[15].PositionInterlock_APLC_Input[1].EquipmentInterlock_APLC_Input[1].SignalInterlock_APLC_Input[1] := "Get Sinais de Interlock Main line".Station[9]."Sinal do job"[0] AND NOT "BYPASS_MOD_2" AND NOT "BYPASS_GERAL" AND NOT "BYPASS_POSTO_QG";
   "Signals".ProcessInterlock_APLC_Input[1].ModezoneInterlock_APLC_Input[2].StationInterlock_APLC_Input[15].PositionInterlock_APLC_Input[1].EquipmentInterlock_APLC_Input[1].SignalInterlock_APLC_Input[2] := "Get Sinais de Interlock Main line".Station[9]."Sinal do job"[1] AND NOT "BYPASS_MOD_2" AND NOT "BYPASS_GERAL" AND NOT "BYPASS_POSTO_QG";
   "Signals".ProcessInterlock_APLC_Input[1].ModezoneInterlock_APLC_Input[2].StationInterlock_APLC_Input[15].PositionInterlock_APLC_Input[1].EquipmentInterlock_APLC_Input[1].SignalInterlock_APLC_Input[3] := NOT "Get Sinais de Interlock Main line".Station[9]."Sinal do job"[2] AND NOT "BYPASS_MOD_2" AND NOT "BYPASS_GERAL" AND NOT "Get Sinais de Interlock Main line".Station[9]."Sinal do job"[9] AND NOT "Get Sinais de Interlock Main line".Station[9]."Sinal do job"[3] AND NOT "Get Sinais de Interlock Main line".Station[9]."Sinal do job"[4] AND NOT "BYPASS_POSTO_QG" AND NOT "Get_Cabine"."SIGNAL RESERVED"[2].BOOL_2 AND NOT "Get_Cabine"."SIGNAL RESERVED"[2].BOOL_3;
   "Signals".ProcessInterlock_APLC_Input[1].ModezoneInterlock_APLC_Input[2].StationInterlock_APLC_Input[15].PositionInterlock_APLC_Input[1].EquipmentInterlock_APLC_Input[2].SignalInterlock_APLC_Input[1] := "Get Sinais de Interlock Main line".Station[9]."Sinal do job"[3] AND NOT "BYPASS_MOD_2" AND NOT "BYPASS_GERAL" AND NOT "BYPASS_POSTO_QG";
   "Signals".ProcessInterlock_APLC_Input[1].ModezoneInterlock_APLC_Input[2].StationInterlock_APLC_Input[15].PositionInterlock_APLC_Input[1].EquipmentInterlock_APLC_Input[2].SignalInterlock_APLC_Input[2] := "Get Sinais de Interlock Main line".Station[9]."Sinal do job"[4] AND NOT "BYPASS_MOD_2" AND NOT "BYPASS_GERAL" AND NOT "BYPASS_POSTO_QG";
   "Signals".ProcessInterlock_APLC_Input[1].ModezoneInterlock_APLC_Input[2].StationInterlock_APLC_Input[15].PositionInterlock_APLC_Input[1].EquipmentInterlock_APLC_Input[1].SignalInterlock_APLC_Input[4] := NOT "Get Sinais de Interlock Main line".Station[10]."Sinal do job"[0] AND NOT "BYPASS_MOD_2" AND NOT "BYPASS_GERAL" AND NOT "BYPASS_POSTO_QG";
   "Signals".ProcessInterlock_APLC_Input[1].ModezoneInterlock_APLC_Input[2].StationInterlock_APLC_Input[15].PositionInterlock_APLC_Input[1].EquipmentInterlock_APLC_Input[2].SignalInterlock_APLC_Input[3] := "GAP_E_EIXO_PENDURADO" AND NOT "BYPASS_MOD_2" AND NOT "BYPASS_GERAL" AND NOT "BYPASS_POSTO_QG";
   "Signals".ProcessInterlock_APLC_Input[1].ModezoneInterlock_APLC_Input[2].StationInterlock_APLC_Input[15].PositionInterlock_APLC_Input[1].EquipmentInterlock_APLC_Input[1].SignalInterlock_APLC_Input[5] := NOT "AREA_TaktTime.SIMPLE_INTERFACE_TAKTTIME_INPUT".TaktTimeWorkhop_APLC_Out[1].TaktTimeProcess_APLC_Out[1].TaktTimeModeZone_APLC_Out[1].Cycle_Done AND ("AREA_TaktTime.INTERFACE_TAKTTIME_INPUT".TaktTimeWorkhop_SPLC_Out[1].TaktTimeProcess_SPLC_Out[1].TaktTimeModeZone_SPLC_Out[1]."Timer" <= T#1S) AND NOT "BYPASS_POSTO_QG";
END_REGION

REGION Network 30: CABINE DEPINTURA
   // ANDON
   // EMERGÊNCIA
   // PORTAS DA CABINE 
   // SINAL OK DO ROBO (SINAL INFORMANDO QUE A PINTURA FOI CONCLUIDA)
   // TALHA FORA DE POSIÇÃO
   // CABINE NOK (INFORMA QUE TEM ALGUMA FALHA NA CABINE)
   // CONFIRMAÇÃO DE RECEITA
   // TAKT LOCAL
   // SIGNAL RESERVED [1] [BOOL ] = ANDON EXPEDIÇÃO
   // SIGNAL RESERVED [1] [BOOL 1] = ESVAZIAMENTO DE LINHA CABINE
   // SIGNAL RESERVED [1] [BOOL 2] = PLATAFORMA
   // SIGNAL RESERVED [1] [BOOL 3] = ANDON CARGA PLATAFORMA
   // SIGNAL RESERVED [2] [BOOL ] = CABINE GIRANDO
   // SIGNAL RESERVED [2] [BOOL 1 ] = SENSOR DE COLISÃO EXPEDIÇÃO
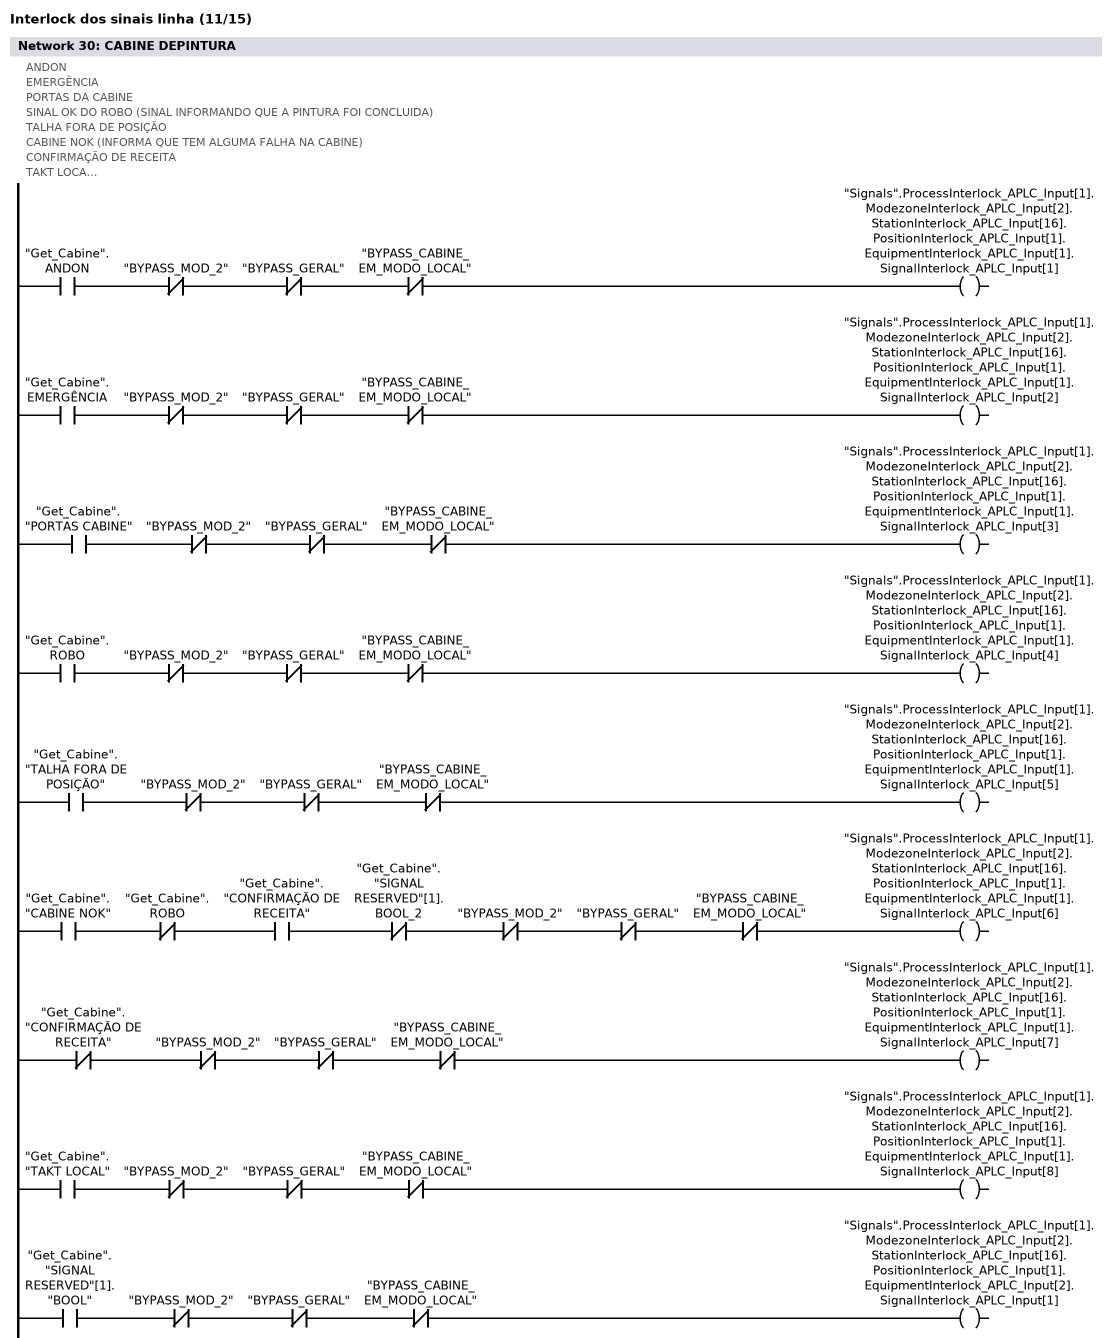
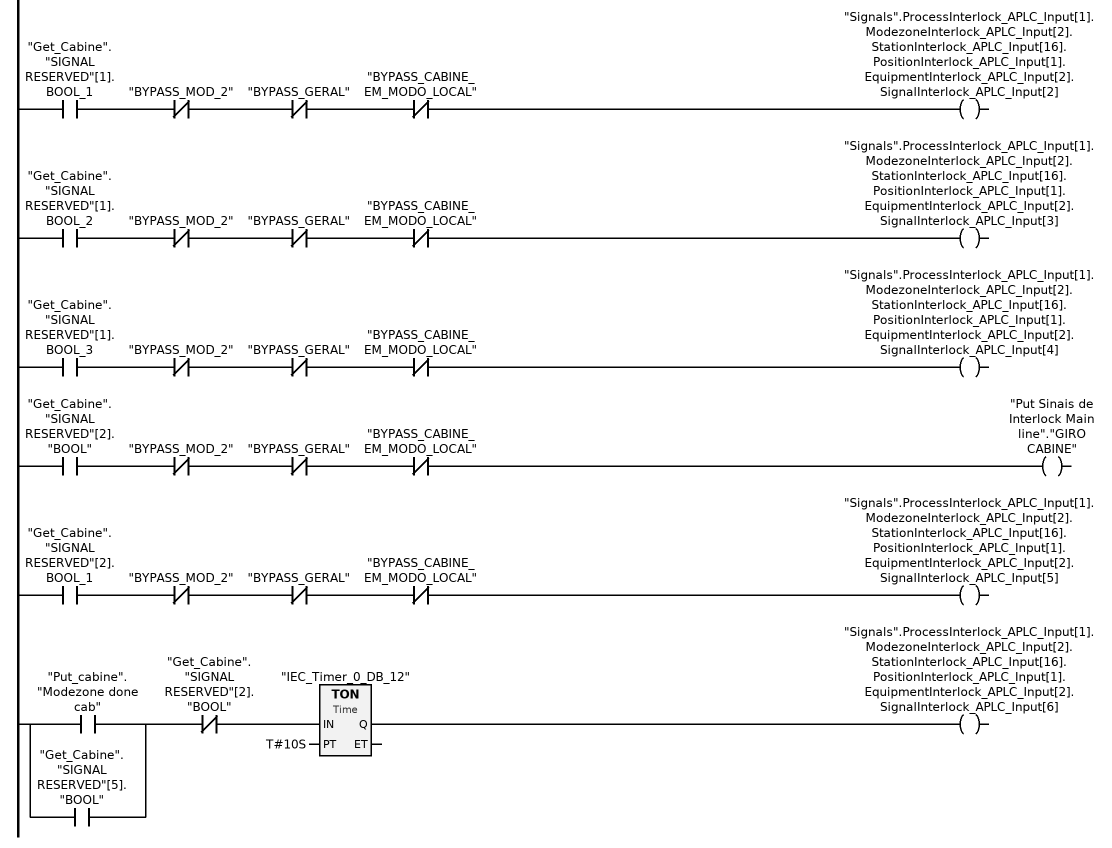
   RUNG wire#powerrail
      Contact( "Get_Cabine".ANDON )
      I_Contact( "BYPASS_MOD_2" )
      I_Contact( "BYPASS_GERAL" )
      I_Contact( "BYPASS_CABINE_EM_MODO_LOCAL" )
      Coil( "Signals".ProcessInterlock_APLC_Input[1].ModezoneInterlock_APLC_Input[2].StationInterlock_APLC_Input[16].PositionInterlock_APLC_Input[1].EquipmentInterlock_APLC_Input[1].SignalInterlock_APLC_Input[1] )
   END_RUNG
   RUNG wire#powerrail
      Contact( "Get_Cabine".EMERGÊNCIA )
      I_Contact( "BYPASS_MOD_2" )
      I_Contact( "BYPASS_GERAL" )
      I_Contact( "BYPASS_CABINE_EM_MODO_LOCAL" )
      Coil( "Signals".ProcessInterlock_APLC_Input[1].ModezoneInterlock_APLC_Input[2].StationInterlock_APLC_Input[16].PositionInterlock_APLC_Input[1].EquipmentInterlock_APLC_Input[1].SignalInterlock_APLC_Input[2] )
   END_RUNG
   RUNG wire#powerrail
      Contact( "Get_Cabine"."PORTAS CABINE" )
      I_Contact( "BYPASS_MOD_2" )
      I_Contact( "BYPASS_GERAL" )
      I_Contact( "BYPASS_CABINE_EM_MODO_LOCAL" )
      Coil( "Signals".ProcessInterlock_APLC_Input[1].ModezoneInterlock_APLC_Input[2].StationInterlock_APLC_Input[16].PositionInterlock_APLC_Input[1].EquipmentInterlock_APLC_Input[1].SignalInterlock_APLC_Input[3] )
   END_RUNG
   RUNG wire#powerrail
      Contact( "Get_Cabine".ROBO )
      I_Contact( "BYPASS_MOD_2" )
      I_Contact( "BYPASS_GERAL" )
      I_Contact( "BYPASS_CABINE_EM_MODO_LOCAL" )
      Coil( "Signals".ProcessInterlock_APLC_Input[1].ModezoneInterlock_APLC_Input[2].StationInterlock_APLC_Input[16].PositionInterlock_APLC_Input[1].EquipmentInterlock_APLC_Input[1].SignalInterlock_APLC_Input[4] )
   END_RUNG
   RUNG wire#powerrail
      Contact( "Get_Cabine"."TALHA FORA DE POSIÇÃO" )
      I_Contact( "BYPASS_MOD_2" )
      I_Contact( "BYPASS_GERAL" )
      I_Contact( "BYPASS_CABINE_EM_MODO_LOCAL" )
      Coil( "Signals".ProcessInterlock_APLC_Input[1].ModezoneInterlock_APLC_Input[2].StationInterlock_APLC_Input[16].PositionInterlock_APLC_Input[1].EquipmentInterlock_APLC_Input[1].SignalInterlock_APLC_Input[5] )
   END_RUNG
   RUNG wire#powerrail
      Contact( "Get_Cabine"."CABINE NOK" )
      I_Contact( "Get_Cabine".ROBO )
      Contact( "Get_Cabine"."CONFIRMAÇÃO DE RECEITA" )
      I_Contact( "Get_Cabine"."SIGNAL RESERVED"[1].BOOL_2 )
      I_Contact( "BYPASS_MOD_2" )
      I_Contact( "BYPASS_GERAL" )
      I_Contact( "BYPASS_CABINE_EM_MODO_LOCAL" )
      Coil( "Signals".ProcessInterlock_APLC_Input[1].ModezoneInterlock_APLC_Input[2].StationInterlock_APLC_Input[16].PositionInterlock_APLC_Input[1].EquipmentInterlock_APLC_Input[1].SignalInterlock_APLC_Input[6] )
   END_RUNG
   RUNG wire#powerrail
      I_Contact( "Get_Cabine"."CONFIRMAÇÃO DE RECEITA" )
      I_Contact( "BYPASS_MOD_2" )
      I_Contact( "BYPASS_GERAL" )
      I_Contact( "BYPASS_CABINE_EM_MODO_LOCAL" )
      Coil( "Signals".ProcessInterlock_APLC_Input[1].ModezoneInterlock_APLC_Input[2].StationInterlock_APLC_Input[16].PositionInterlock_APLC_Input[1].EquipmentInterlock_APLC_Input[1].SignalInterlock_APLC_Input[7] )
   END_RUNG
   RUNG wire#powerrail
      Contact( "Get_Cabine"."TAKT LOCAL" )
      I_Contact( "BYPASS_MOD_2" )
      I_Contact( "BYPASS_GERAL" )
      I_Contact( "BYPASS_CABINE_EM_MODO_LOCAL" )
      Coil( "Signals".ProcessInterlock_APLC_Input[1].ModezoneInterlock_APLC_Input[2].StationInterlock_APLC_Input[16].PositionInterlock_APLC_Input[1].EquipmentInterlock_APLC_Input[1].SignalInterlock_APLC_Input[8] )
   END_RUNG
   RUNG wire#powerrail
      Contact( "Get_Cabine"."SIGNAL RESERVED"[1]."BOOL" )
      I_Contact( "BYPASS_MOD_2" )
      I_Contact( "BYPASS_GERAL" )
      I_Contact( "BYPASS_CABINE_EM_MODO_LOCAL" )
      Coil( "Signals".ProcessInterlock_APLC_Input[1].ModezoneInterlock_APLC_Input[2].StationInterlock_APLC_Input[16].PositionInterlock_APLC_Input[1].EquipmentInterlock_APLC_Input[2].SignalInterlock_APLC_Input[1] )
   END_RUNG
   RUNG wire#powerrail
      Contact( "Get_Cabine"."SIGNAL RESERVED"[1].BOOL_1 )
      I_Contact( "BYPASS_MOD_2" )
      I_Contact( "BYPASS_GERAL" )
      I_Contact( "BYPASS_CABINE_EM_MODO_LOCAL" )
      Coil( "Signals".ProcessInterlock_APLC_Input[1].ModezoneInterlock_APLC_Input[2].StationInterlock_APLC_Input[16].PositionInterlock_APLC_Input[1].EquipmentInterlock_APLC_Input[2].SignalInterlock_APLC_Input[2] )
   END_RUNG
   RUNG wire#powerrail
      Contact( "Get_Cabine"."SIGNAL RESERVED"[1].BOOL_2 )
      I_Contact( "BYPASS_MOD_2" )
      I_Contact( "BYPASS_GERAL" )
      I_Contact( "BYPASS_CABINE_EM_MODO_LOCAL" )
      Coil( "Signals".ProcessInterlock_APLC_Input[1].ModezoneInterlock_APLC_Input[2].StationInterlock_APLC_Input[16].PositionInterlock_APLC_Input[1].EquipmentInterlock_APLC_Input[2].SignalInterlock_APLC_Input[3] )
   END_RUNG
   RUNG wire#powerrail
      Contact( "Get_Cabine"."SIGNAL RESERVED"[1].BOOL_3 )
      I_Contact( "BYPASS_MOD_2" )
      I_Contact( "BYPASS_GERAL" )
      I_Contact( "BYPASS_CABINE_EM_MODO_LOCAL" )
      Coil( "Signals".ProcessInterlock_APLC_Input[1].ModezoneInterlock_APLC_Input[2].StationInterlock_APLC_Input[16].PositionInterlock_APLC_Input[1].EquipmentInterlock_APLC_Input[2].SignalInterlock_APLC_Input[4] )
   END_RUNG
   RUNG wire#powerrail
      Contact( "Get_Cabine"."SIGNAL RESERVED"[2]."BOOL" )
      I_Contact( "BYPASS_MOD_2" )
      I_Contact( "BYPASS_GERAL" )
      I_Contact( "BYPASS_CABINE_EM_MODO_LOCAL" )
      Coil( "Put Sinais de Interlock Main line"."GIRO CABINE" )
   END_RUNG
   RUNG wire#powerrail
      Contact( "Get_Cabine"."SIGNAL RESERVED"[2].BOOL_1 )
      I_Contact( "BYPASS_MOD_2" )
      I_Contact( "BYPASS_GERAL" )
      I_Contact( "BYPASS_CABINE_EM_MODO_LOCAL" )
      Coil( "Signals".ProcessInterlock_APLC_Input[1].ModezoneInterlock_APLC_Input[2].StationInterlock_APLC_Input[16].PositionInterlock_APLC_Input[1].EquipmentInterlock_APLC_Input[2].SignalInterlock_APLC_Input[5] )
   END_RUNG
   RUNG wire#powerrail
      Contact( "Put_cabine"."Modezone done cab" )
      wire#w1
      I_Contact( "Get_Cabine"."SIGNAL RESERVED"[2]."BOOL" )
      { S7_Templates := "time_type := Time" } "IEC_Timer_0_DB_12".TON(pt := T#10S, et =>)
      Coil( "Signals".ProcessInterlock_APLC_Input[1].ModezoneInterlock_APLC_Input[2].StationInterlock_APLC_Input[16].PositionInterlock_APLC_Input[1].EquipmentInterlock_APLC_Input[2].SignalInterlock_APLC_Input[6] )
   END_RUNG
   RUNG wire#powerrail
      Contact( "Get_Cabine"."SIGNAL RESERVED"[5]."BOOL" )
   END_RUNG wire#w1
   // the same network as SCL:
   "Signals".ProcessInterlock_APLC_Input[1].ModezoneInterlock_APLC_Input[2].StationInterlock_APLC_Input[16].PositionInterlock_APLC_Input[1].EquipmentInterlock_APLC_Input[1].SignalInterlock_APLC_Input[1] := "Get_Cabine".ANDON AND NOT "BYPASS_MOD_2" AND NOT "BYPASS_GERAL" AND NOT "BYPASS_CABINE_EM_MODO_LOCAL";
   "Signals".ProcessInterlock_APLC_Input[1].ModezoneInterlock_APLC_Input[2].StationInterlock_APLC_Input[16].PositionInterlock_APLC_Input[1].EquipmentInterlock_APLC_Input[1].SignalInterlock_APLC_Input[2] := "Get_Cabine".EMERGÊNCIA AND NOT "BYPASS_MOD_2" AND NOT "BYPASS_GERAL" AND NOT "BYPASS_CABINE_EM_MODO_LOCAL";
   "Signals".ProcessInterlock_APLC_Input[1].ModezoneInterlock_APLC_Input[2].StationInterlock_APLC_Input[16].PositionInterlock_APLC_Input[1].EquipmentInterlock_APLC_Input[1].SignalInterlock_APLC_Input[3] := "Get_Cabine"."PORTAS CABINE" AND NOT "BYPASS_MOD_2" AND NOT "BYPASS_GERAL" AND NOT "BYPASS_CABINE_EM_MODO_LOCAL";
   "Signals".ProcessInterlock_APLC_Input[1].ModezoneInterlock_APLC_Input[2].StationInterlock_APLC_Input[16].PositionInterlock_APLC_Input[1].EquipmentInterlock_APLC_Input[1].SignalInterlock_APLC_Input[4] := "Get_Cabine".ROBO AND NOT "BYPASS_MOD_2" AND NOT "BYPASS_GERAL" AND NOT "BYPASS_CABINE_EM_MODO_LOCAL";
   "Signals".ProcessInterlock_APLC_Input[1].ModezoneInterlock_APLC_Input[2].StationInterlock_APLC_Input[16].PositionInterlock_APLC_Input[1].EquipmentInterlock_APLC_Input[1].SignalInterlock_APLC_Input[5] := "Get_Cabine"."TALHA FORA DE POSIÇÃO" AND NOT "BYPASS_MOD_2" AND NOT "BYPASS_GERAL" AND NOT "BYPASS_CABINE_EM_MODO_LOCAL";
   "Signals".ProcessInterlock_APLC_Input[1].ModezoneInterlock_APLC_Input[2].StationInterlock_APLC_Input[16].PositionInterlock_APLC_Input[1].EquipmentInterlock_APLC_Input[1].SignalInterlock_APLC_Input[6] := "Get_Cabine"."CABINE NOK" AND NOT "Get_Cabine".ROBO AND "Get_Cabine"."CONFIRMAÇÃO DE RECEITA" AND NOT "Get_Cabine"."SIGNAL RESERVED"[1].BOOL_2 AND NOT "BYPASS_MOD_2" AND NOT "BYPASS_GERAL" AND NOT "BYPASS_CABINE_EM_MODO_LOCAL";
   "Signals".ProcessInterlock_APLC_Input[1].ModezoneInterlock_APLC_Input[2].StationInterlock_APLC_Input[16].PositionInterlock_APLC_Input[1].EquipmentInterlock_APLC_Input[1].SignalInterlock_APLC_Input[7] := NOT "Get_Cabine"."CONFIRMAÇÃO DE RECEITA" AND NOT "BYPASS_MOD_2" AND NOT "BYPASS_GERAL" AND NOT "BYPASS_CABINE_EM_MODO_LOCAL";
   "Signals".ProcessInterlock_APLC_Input[1].ModezoneInterlock_APLC_Input[2].StationInterlock_APLC_Input[16].PositionInterlock_APLC_Input[1].EquipmentInterlock_APLC_Input[1].SignalInterlock_APLC_Input[8] := "Get_Cabine"."TAKT LOCAL" AND NOT "BYPASS_MOD_2" AND NOT "BYPASS_GERAL" AND NOT "BYPASS_CABINE_EM_MODO_LOCAL";
   "Signals".ProcessInterlock_APLC_Input[1].ModezoneInterlock_APLC_Input[2].StationInterlock_APLC_Input[16].PositionInterlock_APLC_Input[1].EquipmentInterlock_APLC_Input[2].SignalInterlock_APLC_Input[1] := "Get_Cabine"."SIGNAL RESERVED"[1]."BOOL" AND NOT "BYPASS_MOD_2" AND NOT "BYPASS_GERAL" AND NOT "BYPASS_CABINE_EM_MODO_LOCAL";
   "Signals".ProcessInterlock_APLC_Input[1].ModezoneInterlock_APLC_Input[2].StationInterlock_APLC_Input[16].PositionInterlock_APLC_Input[1].EquipmentInterlock_APLC_Input[2].SignalInterlock_APLC_Input[2] := "Get_Cabine"."SIGNAL RESERVED"[1].BOOL_1 AND NOT "BYPASS_MOD_2" AND NOT "BYPASS_GERAL" AND NOT "BYPASS_CABINE_EM_MODO_LOCAL";
   "Signals".ProcessInterlock_APLC_Input[1].ModezoneInterlock_APLC_Input[2].StationInterlock_APLC_Input[16].PositionInterlock_APLC_Input[1].EquipmentInterlock_APLC_Input[2].SignalInterlock_APLC_Input[3] := "Get_Cabine"."SIGNAL RESERVED"[1].BOOL_2 AND NOT "BYPASS_MOD_2" AND NOT "BYPASS_GERAL" AND NOT "BYPASS_CABINE_EM_MODO_LOCAL";
   "Signals".ProcessInterlock_APLC_Input[1].ModezoneInterlock_APLC_Input[2].StationInterlock_APLC_Input[16].PositionInterlock_APLC_Input[1].EquipmentInterlock_APLC_Input[2].SignalInterlock_APLC_Input[4] := "Get_Cabine"."SIGNAL RESERVED"[1].BOOL_3 AND NOT "BYPASS_MOD_2" AND NOT "BYPASS_GERAL" AND NOT "BYPASS_CABINE_EM_MODO_LOCAL";
   "Put Sinais de Interlock Main line"."GIRO CABINE" := "Get_Cabine"."SIGNAL RESERVED"[2]."BOOL" AND NOT "BYPASS_MOD_2" AND NOT "BYPASS_GERAL" AND NOT "BYPASS_CABINE_EM_MODO_LOCAL";
   "Signals".ProcessInterlock_APLC_Input[1].ModezoneInterlock_APLC_Input[2].StationInterlock_APLC_Input[16].PositionInterlock_APLC_Input[1].EquipmentInterlock_APLC_Input[2].SignalInterlock_APLC_Input[5] := "Get_Cabine"."SIGNAL RESERVED"[2].BOOL_1 AND NOT "BYPASS_MOD_2" AND NOT "BYPASS_GERAL" AND NOT "BYPASS_CABINE_EM_MODO_LOCAL";
   "IEC_Timer_0_DB_12".TON(IN := ("Put_cabine"."Modezone done cab" OR "Get_Cabine"."SIGNAL RESERVED"[5]."BOOL") AND NOT "Get_Cabine"."SIGNAL RESERVED"[2]."BOOL",
                           PT := T#10S);
   "Signals".ProcessInterlock_APLC_Input[1].ModezoneInterlock_APLC_Input[2].StationInterlock_APLC_Input[16].PositionInterlock_APLC_Input[1].EquipmentInterlock_APLC_Input[2].SignalInterlock_APLC_Input[6] := "IEC_Timer_0_DB_12".Q;
END_REGION

REGION Network 31: SINAIS ENVIADOS PARA CABINE
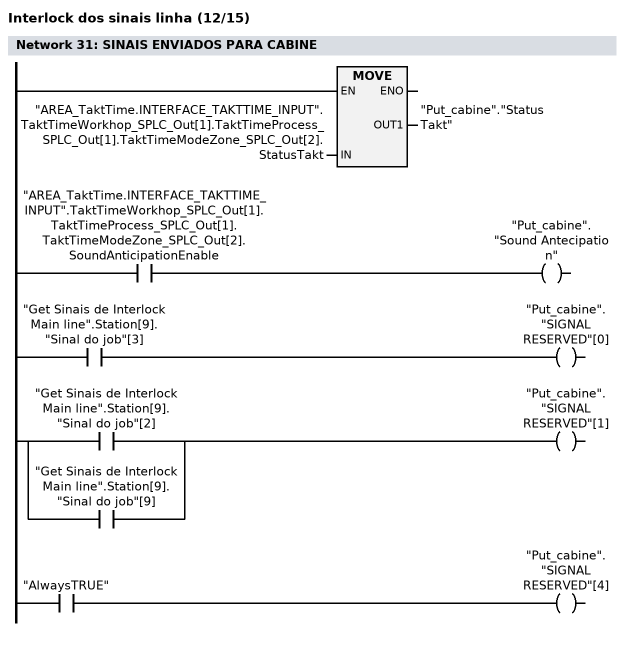
   RUNG wire#powerrail
      Move(in := "AREA_TaktTime.INTERFACE_TAKTTIME_INPUT".TaktTimeWorkhop_SPLC_Out[1].TaktTimeProcess_SPLC_Out[1].TaktTimeModeZone_SPLC_Out[2].StatusTakt, out1 => "Put_cabine"."Status Takt")
   END_RUNG
   RUNG wire#powerrail
      Contact( "AREA_TaktTime.INTERFACE_TAKTTIME_INPUT".TaktTimeWorkhop_SPLC_Out[1].TaktTimeProcess_SPLC_Out[1].TaktTimeModeZone_SPLC_Out[2].SoundAnticipationEnable )
      Coil( "Put_cabine"."Sound Antecipation" )
   END_RUNG
   RUNG wire#powerrail
      Contact( "Get Sinais de Interlock Main line".Station[9]."Sinal do job"[3] )
      Coil( "Put_cabine"."SIGNAL RESERVED"[0] )
   END_RUNG
   RUNG wire#powerrail
      Contact( "Get Sinais de Interlock Main line".Station[9]."Sinal do job"[2] )
      wire#w1
      Coil( "Put_cabine"."SIGNAL RESERVED"[1] )
   END_RUNG
   RUNG wire#powerrail
      Contact( "Get Sinais de Interlock Main line".Station[9]."Sinal do job"[9] )
   END_RUNG wire#w1
   RUNG wire#powerrail
      Contact( "AlwaysTRUE" )
      Coil( "Put_cabine"."SIGNAL RESERVED"[4] )
   END_RUNG
   // the same network as SCL:
   "Put_cabine"."Status Takt" := "AREA_TaktTime.INTERFACE_TAKTTIME_INPUT".TaktTimeWorkhop_SPLC_Out[1].TaktTimeProcess_SPLC_Out[1].TaktTimeModeZone_SPLC_Out[2].StatusTakt;
   "Put_cabine"."Sound Antecipation" := "AREA_TaktTime.INTERFACE_TAKTTIME_INPUT".TaktTimeWorkhop_SPLC_Out[1].TaktTimeProcess_SPLC_Out[1].TaktTimeModeZone_SPLC_Out[2].SoundAnticipationEnable;
   "Put_cabine"."SIGNAL RESERVED"[0] := "Get Sinais de Interlock Main line".Station[9]."Sinal do job"[3];
   "Put_cabine"."SIGNAL RESERVED"[1] := "Get Sinais de Interlock Main line".Station[9]."Sinal do job"[2] OR "Get Sinais de Interlock Main line".Station[9]."Sinal do job"[9];
   "Put_cabine"."SIGNAL RESERVED"[4] := "AlwaysTRUE";
END_REGION

REGION Network 32: Mod1 e 2 OK
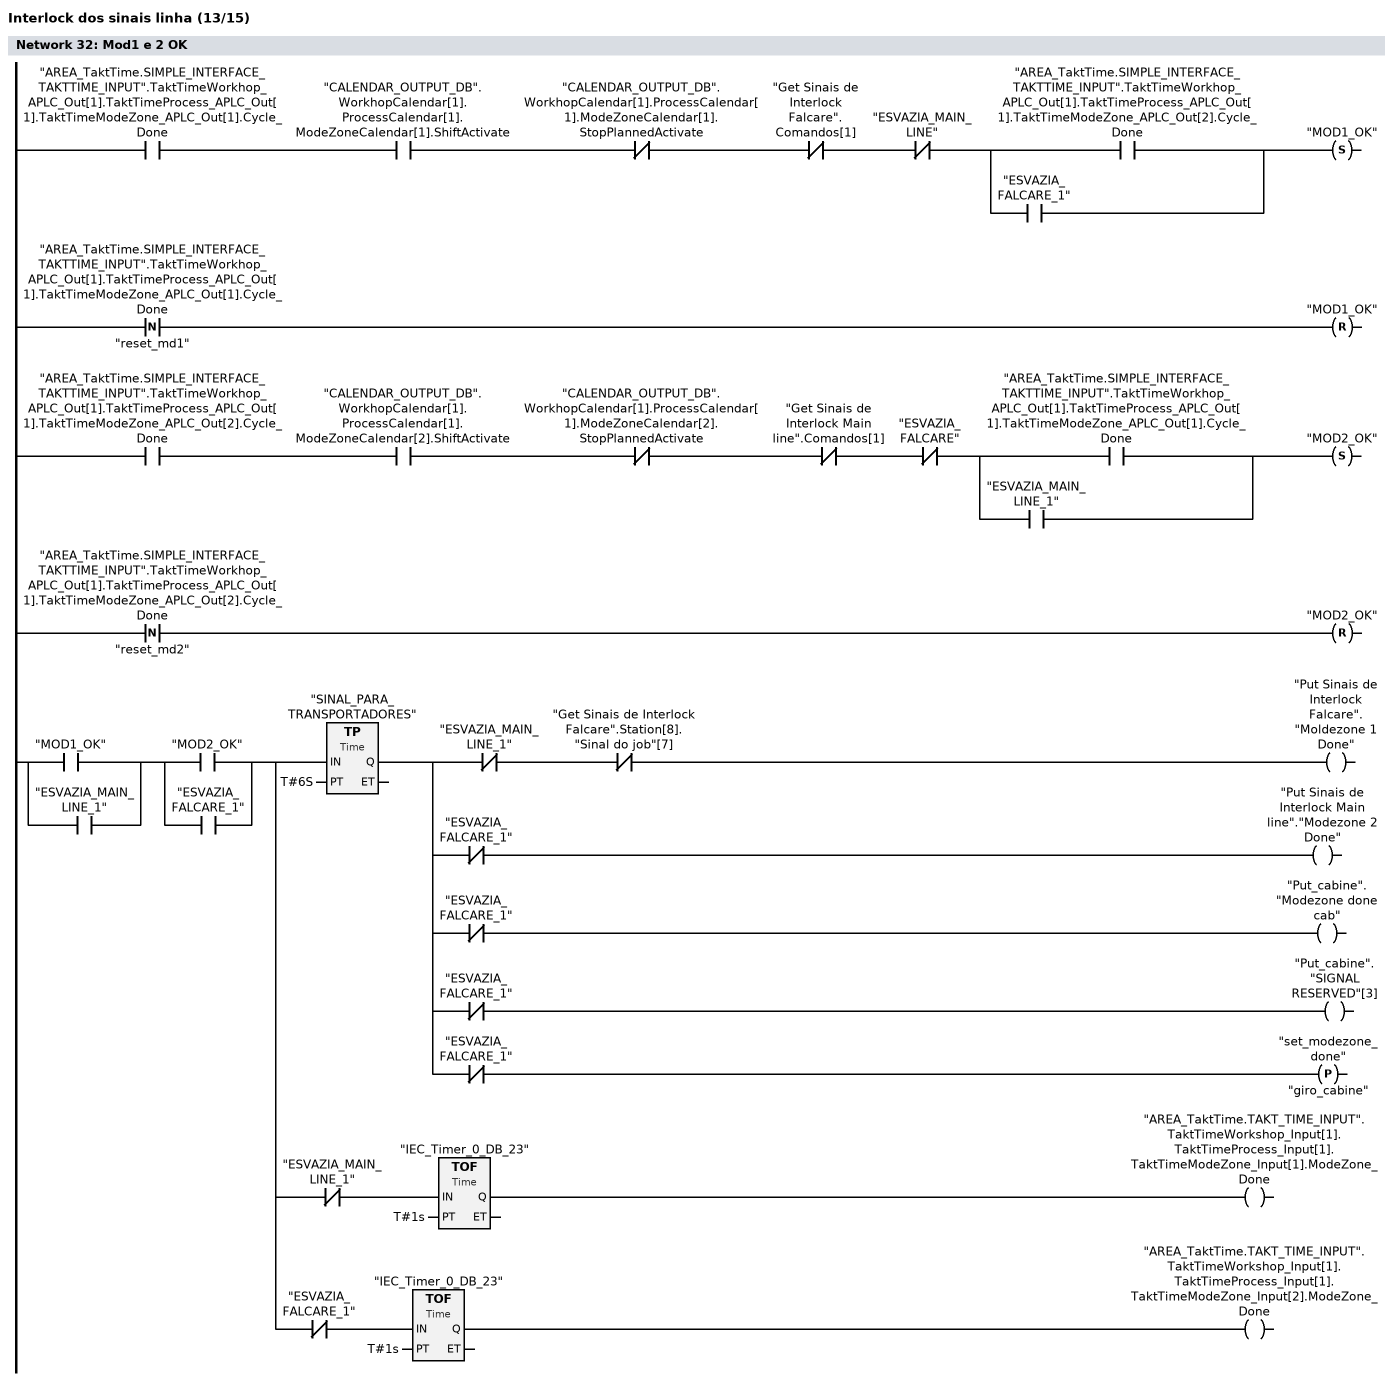
   IF "AREA_TaktTime.SIMPLE_INTERFACE_TAKTTIME_INPUT".TaktTimeWorkhop_APLC_Out[1].TaktTimeProcess_APLC_Out[1].TaktTimeModeZone_APLC_Out[1].Cycle_Done AND "CALENDAR_OUTPUT_DB".WorkhopCalendar[1].ProcessCalendar[1].ModeZoneCalendar[1].ShiftActivate AND NOT "CALENDAR_OUTPUT_DB".WorkhopCalendar[1].ProcessCalendar[1].ModeZoneCalendar[1].StopPlannedActivate AND NOT "Get Sinais de Interlock Falcare".Comandos[1] AND NOT "ESVAZIA_MAIN_LINE" AND ("AREA_TaktTime.SIMPLE_INTERFACE_TAKTTIME_INPUT".TaktTimeWorkhop_APLC_Out[1].TaktTimeProcess_APLC_Out[1].TaktTimeModeZone_APLC_Out[2].Cycle_Done OR "ESVAZIA_FALCARE_1") THEN
       "MOD1_OK" := TRUE;
   END_IF;
   #_w1 := NOT "AREA_TaktTime.SIMPLE_INTERFACE_TAKTTIME_INPUT".TaktTimeWorkhop_APLC_Out[1].TaktTimeProcess_APLC_Out[1].TaktTimeModeZone_APLC_Out[1].Cycle_Done AND "reset_md1";   // falling edge of "AREA_TaktTime.SIMPLE_INTERFACE_TAKTTIME_INPUT".TaktTimeWorkhop_APLC_Out[1].TaktTimeProcess_APLC_Out[1].TaktTimeModeZone_APLC_Out[1].Cycle_Done
   "reset_md1" := "AREA_TaktTime.SIMPLE_INTERFACE_TAKTTIME_INPUT".TaktTimeWorkhop_APLC_Out[1].TaktTimeProcess_APLC_Out[1].TaktTimeModeZone_APLC_Out[1].Cycle_Done;
   IF #_w1 THEN "MOD1_OK" := FALSE; END_IF;
   IF "AREA_TaktTime.SIMPLE_INTERFACE_TAKTTIME_INPUT".TaktTimeWorkhop_APLC_Out[1].TaktTimeProcess_APLC_Out[1].TaktTimeModeZone_APLC_Out[2].Cycle_Done AND "CALENDAR_OUTPUT_DB".WorkhopCalendar[1].ProcessCalendar[1].ModeZoneCalendar[2].ShiftActivate AND NOT "CALENDAR_OUTPUT_DB".WorkhopCalendar[1].ProcessCalendar[1].ModeZoneCalendar[2].StopPlannedActivate AND NOT "Get Sinais de Interlock Main line".Comandos[1] AND NOT "ESVAZIA_FALCARE" AND ("AREA_TaktTime.SIMPLE_INTERFACE_TAKTTIME_INPUT".TaktTimeWorkhop_APLC_Out[1].TaktTimeProcess_APLC_Out[1].TaktTimeModeZone_APLC_Out[1].Cycle_Done OR "ESVAZIA_MAIN_LINE_1") THEN
       "MOD2_OK" := TRUE;
   END_IF;
   #_w2 := NOT "AREA_TaktTime.SIMPLE_INTERFACE_TAKTTIME_INPUT".TaktTimeWorkhop_APLC_Out[1].TaktTimeProcess_APLC_Out[1].TaktTimeModeZone_APLC_Out[2].Cycle_Done AND "reset_md2";   // falling edge of "AREA_TaktTime.SIMPLE_INTERFACE_TAKTTIME_INPUT".TaktTimeWorkhop_APLC_Out[1].TaktTimeProcess_APLC_Out[1].TaktTimeModeZone_APLC_Out[2].Cycle_Done
   "reset_md2" := "AREA_TaktTime.SIMPLE_INTERFACE_TAKTTIME_INPUT".TaktTimeWorkhop_APLC_Out[1].TaktTimeProcess_APLC_Out[1].TaktTimeModeZone_APLC_Out[2].Cycle_Done;
   IF #_w2 THEN "MOD2_OK" := FALSE; END_IF;
   #_w3 := ("MOD1_OK" OR "ESVAZIA_MAIN_LINE_1") AND ("MOD2_OK" OR "ESVAZIA_FALCARE_1");
   "SINAL_PARA_TRANSPORTADORES".TP(IN := #_w3, PT := T#6S);
   "Put Sinais de Interlock Falcare"."Moldezone 1 Done" := "SINAL_PARA_TRANSPORTADORES".Q AND NOT "ESVAZIA_MAIN_LINE_1" AND NOT "Get Sinais de Interlock Falcare".Station[8]."Sinal do job"[7];
   "Put Sinais de Interlock Main line"."Modezone 2 Done" := "SINAL_PARA_TRANSPORTADORES".Q AND NOT "ESVAZIA_FALCARE_1";
   "Put_cabine"."Modezone done cab" := "SINAL_PARA_TRANSPORTADORES".Q AND NOT "ESVAZIA_FALCARE_1";
   "Put_cabine"."SIGNAL RESERVED"[3] := "SINAL_PARA_TRANSPORTADORES".Q AND NOT "ESVAZIA_FALCARE_1";
   #_w4 := "SINAL_PARA_TRANSPORTADORES".Q AND NOT "ESVAZIA_FALCARE_1";
   "set_modezone_done" := #_w4 AND NOT "giro_cabine";   // rising edge
   "giro_cabine" := #_w4;
   "IEC_Timer_0_DB_23".TOF(IN := #_w3 AND NOT "ESVAZIA_MAIN_LINE_1", PT := T#1s);
   "AREA_TaktTime.TAKT_TIME_INPUT".TaktTimeWorkshop_Input[1].TaktTimeProcess_Input[1].TaktTimeModeZone_Input[1].ModeZone_Done := "IEC_Timer_0_DB_23".Q;
   "IEC_Timer_0_DB_23".TOF(IN := #_w3 AND NOT "ESVAZIA_FALCARE_1", PT := T#1s);
   "AREA_TaktTime.TAKT_TIME_INPUT".TaktTimeWorkshop_Input[1].TaktTimeProcess_Input[1].TaktTimeModeZone_Input[2].ModeZone_Done := "IEC_Timer_0_DB_23".Q;
END_REGION

REGION Network 33: LIBERAÇÃO DE TURNO ATIVO PARA TRANSPORTADORES FALCARE E MAIN LINE / CABINE DE PINTURA
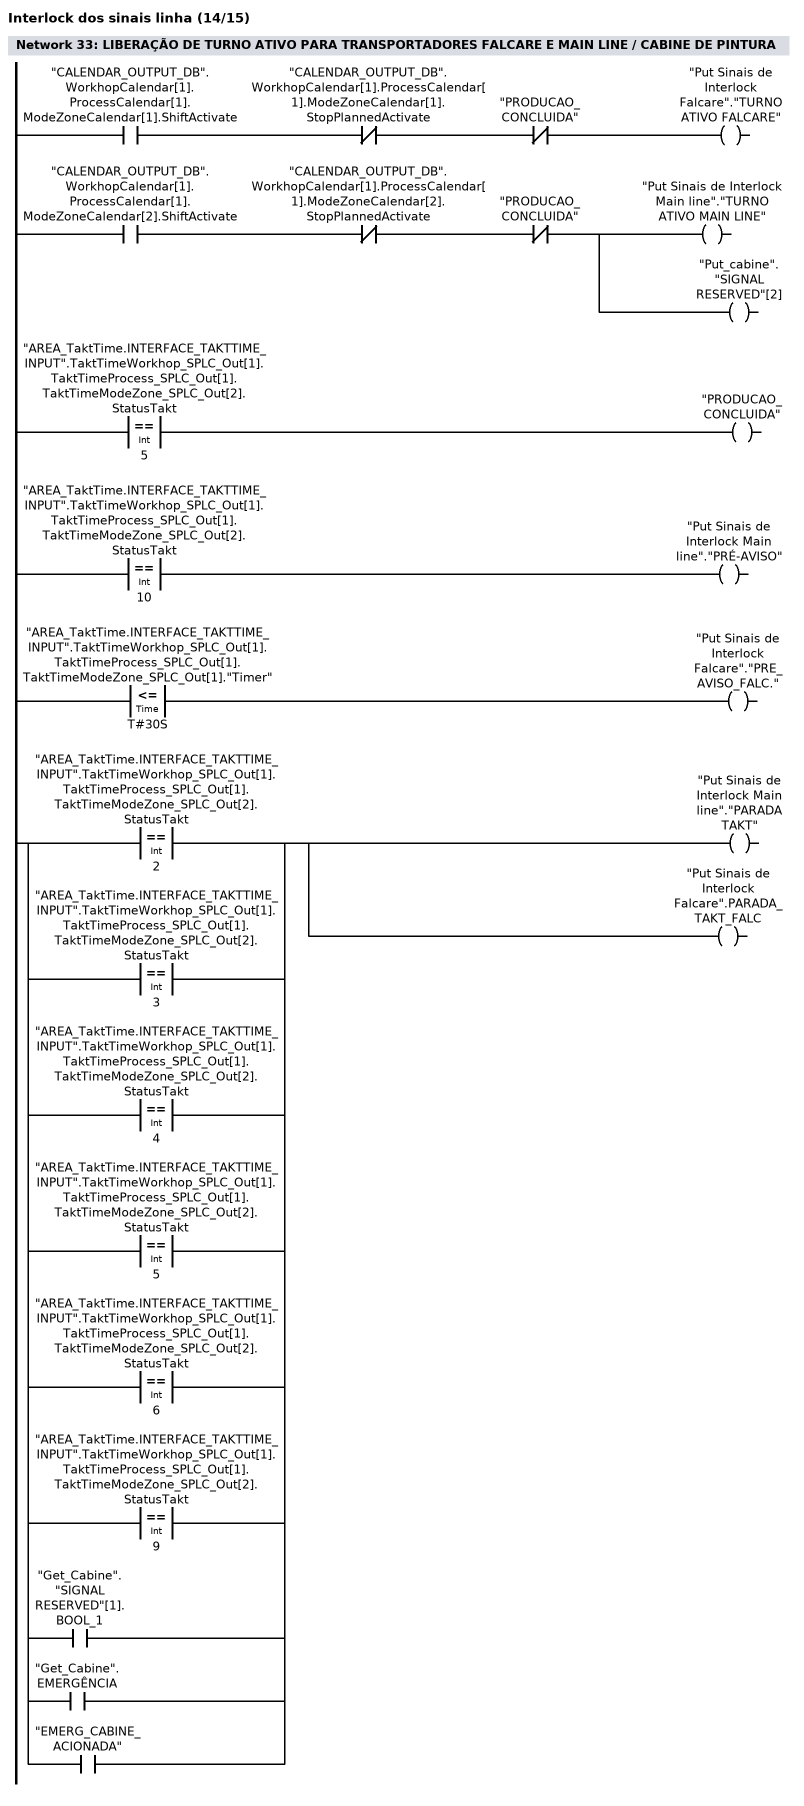
   RUNG wire#powerrail
      Contact( "CALENDAR_OUTPUT_DB".WorkhopCalendar[1].ProcessCalendar[1].ModeZoneCalendar[1].ShiftActivate )
      I_Contact( "CALENDAR_OUTPUT_DB".WorkhopCalendar[1].ProcessCalendar[1].ModeZoneCalendar[1].StopPlannedActivate )
      I_Contact( "PRODUCAO_CONCLUIDA" )
      Coil( "Put Sinais de Interlock Falcare"."TURNO ATIVO FALCARE" )
   END_RUNG
   RUNG wire#powerrail
      Contact( "CALENDAR_OUTPUT_DB".WorkhopCalendar[1].ProcessCalendar[1].ModeZoneCalendar[2].ShiftActivate )
      I_Contact( "CALENDAR_OUTPUT_DB".WorkhopCalendar[1].ProcessCalendar[1].ModeZoneCalendar[2].StopPlannedActivate )
      I_Contact( "PRODUCAO_CONCLUIDA" )
      wire#w1
      Coil( "Put Sinais de Interlock Main line"."TURNO ATIVO MAIN LINE" )
   END_RUNG
   RUNG wire#w1
      Coil( "Put_cabine"."SIGNAL RESERVED"[2] )
   END_RUNG
   RUNG wire#powerrail
      { S7_Templates := "SrcType := Int" } EQ_Contact(in1 := "AREA_TaktTime.INTERFACE_TAKTTIME_INPUT".TaktTimeWorkhop_SPLC_Out[1].TaktTimeProcess_SPLC_Out[1].TaktTimeModeZone_SPLC_Out[2].StatusTakt, in2 := 5)
      Coil( "PRODUCAO_CONCLUIDA" )
   END_RUNG
   RUNG wire#powerrail
      { S7_Templates := "SrcType := Int" } EQ_Contact(in1 := "AREA_TaktTime.INTERFACE_TAKTTIME_INPUT".TaktTimeWorkhop_SPLC_Out[1].TaktTimeProcess_SPLC_Out[1].TaktTimeModeZone_SPLC_Out[2].StatusTakt, in2 := 10)
      Coil( "Put Sinais de Interlock Main line"."PRÉ-AVISO" )
   END_RUNG
   RUNG wire#powerrail
      { S7_Templates := "SrcType := Time" } LE_Contact(in1 := "AREA_TaktTime.INTERFACE_TAKTTIME_INPUT".TaktTimeWorkhop_SPLC_Out[1].TaktTimeProcess_SPLC_Out[1].TaktTimeModeZone_SPLC_Out[1]."Timer", in2 := T#30S)
      Coil( "Put Sinais de Interlock Falcare"."PRE_AVISO_FALC." )
   END_RUNG
   RUNG wire#powerrail
      { S7_Templates := "SrcType := Int" } EQ_Contact(in1 := "AREA_TaktTime.INTERFACE_TAKTTIME_INPUT".TaktTimeWorkhop_SPLC_Out[1].TaktTimeProcess_SPLC_Out[1].TaktTimeModeZone_SPLC_Out[2].StatusTakt, in2 := 2)
      wire#w2
      Coil( "Put Sinais de Interlock Main line"."PARADA TAKT" )
   END_RUNG
   RUNG wire#powerrail
      { S7_Templates := "SrcType := Int" } EQ_Contact(in1 := "AREA_TaktTime.INTERFACE_TAKTTIME_INPUT".TaktTimeWorkhop_SPLC_Out[1].TaktTimeProcess_SPLC_Out[1].TaktTimeModeZone_SPLC_Out[2].StatusTakt, in2 := 3)
   END_RUNG wire#w2
   RUNG wire#powerrail
      { S7_Templates := "SrcType := Int" } EQ_Contact(in1 := "AREA_TaktTime.INTERFACE_TAKTTIME_INPUT".TaktTimeWorkhop_SPLC_Out[1].TaktTimeProcess_SPLC_Out[1].TaktTimeModeZone_SPLC_Out[2].StatusTakt, in2 := 4)
   END_RUNG wire#w2
   RUNG wire#powerrail
      { S7_Templates := "SrcType := Int" } EQ_Contact(in1 := "AREA_TaktTime.INTERFACE_TAKTTIME_INPUT".TaktTimeWorkhop_SPLC_Out[1].TaktTimeProcess_SPLC_Out[1].TaktTimeModeZone_SPLC_Out[2].StatusTakt, in2 := 5)
   END_RUNG wire#w2
   RUNG wire#powerrail
      { S7_Templates := "SrcType := Int" } EQ_Contact(in1 := "AREA_TaktTime.INTERFACE_TAKTTIME_INPUT".TaktTimeWorkhop_SPLC_Out[1].TaktTimeProcess_SPLC_Out[1].TaktTimeModeZone_SPLC_Out[2].StatusTakt, in2 := 6)
   END_RUNG wire#w2
   RUNG wire#powerrail
      { S7_Templates := "SrcType := Int" } EQ_Contact(in1 := "AREA_TaktTime.INTERFACE_TAKTTIME_INPUT".TaktTimeWorkhop_SPLC_Out[1].TaktTimeProcess_SPLC_Out[1].TaktTimeModeZone_SPLC_Out[2].StatusTakt, in2 := 9)
   END_RUNG wire#w2
   RUNG wire#powerrail
      Contact( "Get_Cabine"."SIGNAL RESERVED"[1].BOOL_1 )
   END_RUNG wire#w2
   RUNG wire#powerrail
      Contact( "Get_Cabine".EMERGÊNCIA )
   END_RUNG wire#w2
   RUNG wire#powerrail
      Contact( "EMERG_CABINE_ACIONADA" )
   END_RUNG wire#w2
   RUNG wire#w2
      Coil( "Put Sinais de Interlock Falcare".PARADA_TAKT_FALC )
   END_RUNG
   // the same network as SCL:
   "Put Sinais de Interlock Falcare"."TURNO ATIVO FALCARE" := "CALENDAR_OUTPUT_DB".WorkhopCalendar[1].ProcessCalendar[1].ModeZoneCalendar[1].ShiftActivate AND NOT "CALENDAR_OUTPUT_DB".WorkhopCalendar[1].ProcessCalendar[1].ModeZoneCalendar[1].StopPlannedActivate AND NOT "PRODUCAO_CONCLUIDA";
   "Put Sinais de Interlock Main line"."TURNO ATIVO MAIN LINE" := "CALENDAR_OUTPUT_DB".WorkhopCalendar[1].ProcessCalendar[1].ModeZoneCalendar[2].ShiftActivate AND NOT "CALENDAR_OUTPUT_DB".WorkhopCalendar[1].ProcessCalendar[1].ModeZoneCalendar[2].StopPlannedActivate AND NOT "PRODUCAO_CONCLUIDA";
   "Put_cabine"."SIGNAL RESERVED"[2] := "Put Sinais de Interlock Main line"."TURNO ATIVO MAIN LINE";
   "PRODUCAO_CONCLUIDA" := "AREA_TaktTime.INTERFACE_TAKTTIME_INPUT".TaktTimeWorkhop_SPLC_Out[1].TaktTimeProcess_SPLC_Out[1].TaktTimeModeZone_SPLC_Out[2].StatusTakt = 5;
   "Put Sinais de Interlock Main line"."PRÉ-AVISO" := "AREA_TaktTime.INTERFACE_TAKTTIME_INPUT".TaktTimeWorkhop_SPLC_Out[1].TaktTimeProcess_SPLC_Out[1].TaktTimeModeZone_SPLC_Out[2].StatusTakt = 10;
   "Put Sinais de Interlock Falcare"."PRE_AVISO_FALC." := "AREA_TaktTime.INTERFACE_TAKTTIME_INPUT".TaktTimeWorkhop_SPLC_Out[1].TaktTimeProcess_SPLC_Out[1].TaktTimeModeZone_SPLC_Out[1]."Timer" <= T#30S;
   "Put Sinais de Interlock Main line"."PARADA TAKT" := ("AREA_TaktTime.INTERFACE_TAKTTIME_INPUT".TaktTimeWorkhop_SPLC_Out[1].TaktTimeProcess_SPLC_Out[1].TaktTimeModeZone_SPLC_Out[2].StatusTakt = 2) OR ("AREA_TaktTime.INTERFACE_TAKTTIME_INPUT".TaktTimeWorkhop_SPLC_Out[1].TaktTimeProcess_SPLC_Out[1].TaktTimeModeZone_SPLC_Out[2].StatusTakt = 3) OR ("AREA_TaktTime.INTERFACE_TAKTTIME_INPUT".TaktTimeWorkhop_SPLC_Out[1].TaktTimeProcess_SPLC_Out[1].TaktTimeModeZone_SPLC_Out[2].StatusTakt = 4) OR ("AREA_TaktTime.INTERFACE_TAKTTIME_INPUT".TaktTimeWorkhop_SPLC_Out[1].TaktTimeProcess_SPLC_Out[1].TaktTimeModeZone_SPLC_Out[2].StatusTakt = 5) OR ("AREA_TaktTime.INTERFACE_TAKTTIME_INPUT".TaktTimeWorkhop_SPLC_Out[1].TaktTimeProcess_SPLC_Out[1].TaktTimeModeZone_SPLC_Out[2].StatusTakt = 6) OR ("AREA_TaktTime.INTERFACE_TAKTTIME_INPUT".TaktTimeWorkhop_SPLC_Out[1].TaktTimeProcess_SPLC_Out[1].TaktTimeModeZone_SPLC_Out[2].StatusTakt = 9) OR "Get_Cabine"."SIGNAL RESERVED"[1].BOOL_1 OR "Get_Cabine".EMERGÊNCIA OR "EMERG_CABINE_ACIONADA";
   "Put Sinais de Interlock Falcare".PARADA_TAKT_FALC := "Put Sinais de Interlock Main line"."PARADA TAKT";
END_REGION

REGION Network 34: LIFE BIT PARA TRANSPORTADORES
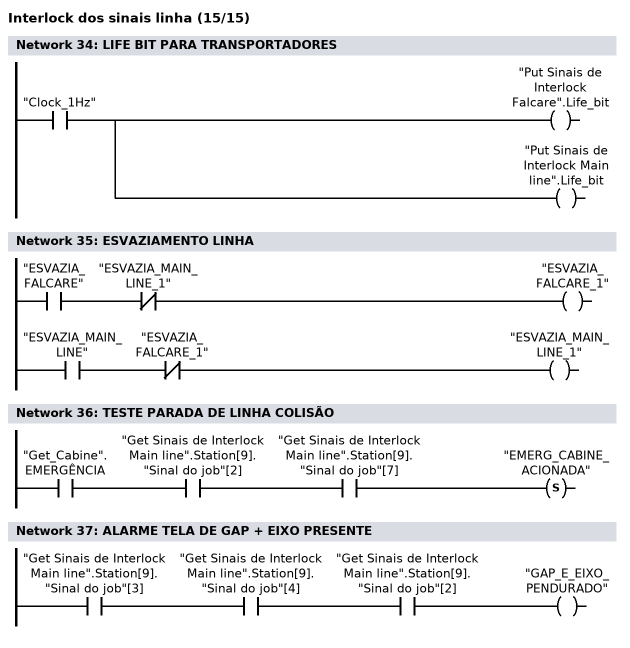
   RUNG wire#powerrail
      Contact( "Clock_1Hz" )
      wire#w1
      Coil( "Put Sinais de Interlock Falcare".Life_bit )
   END_RUNG
   RUNG wire#w1
      Coil( "Put Sinais de Interlock Main line".Life_bit )
   END_RUNG
   // the same network as SCL:
   "Put Sinais de Interlock Falcare".Life_bit := "Clock_1Hz";
   "Put Sinais de Interlock Main line".Life_bit := "Clock_1Hz";
END_REGION

REGION Network 35: ESVAZIAMENTO LINHA
   RUNG wire#powerrail
      Contact( "ESVAZIA_FALCARE" )
      I_Contact( "ESVAZIA_MAIN_LINE_1" )
      Coil( "ESVAZIA_FALCARE_1" )
   END_RUNG
   RUNG wire#powerrail
      Contact( "ESVAZIA_MAIN_LINE" )
      I_Contact( "ESVAZIA_FALCARE_1" )
      Coil( "ESVAZIA_MAIN_LINE_1" )
   END_RUNG
   // the same network as SCL:
   "ESVAZIA_FALCARE_1" := "ESVAZIA_FALCARE" AND NOT "ESVAZIA_MAIN_LINE_1";
   "ESVAZIA_MAIN_LINE_1" := "ESVAZIA_MAIN_LINE" AND NOT "ESVAZIA_FALCARE_1";
END_REGION

REGION Network 36: TESTE PARADA DE LINHA COLISÃO
   RUNG wire#powerrail
      Contact( "Get_Cabine".EMERGÊNCIA )
      Contact( "Get Sinais de Interlock Main line".Station[9]."Sinal do job"[2] )
      Contact( "Get Sinais de Interlock Main line".Station[9]."Sinal do job"[7] )
      S_Coil( "EMERG_CABINE_ACIONADA" )
   END_RUNG
   // the same network as SCL:
   IF "Get_Cabine".EMERGÊNCIA AND "Get Sinais de Interlock Main line".Station[9]."Sinal do job"[2] AND "Get Sinais de Interlock Main line".Station[9]."Sinal do job"[7] THEN
       "EMERG_CABINE_ACIONADA" := TRUE;
   END_IF;
END_REGION

REGION Network 37: ALARME TELA DE GAP + EIXO PRESENTE
   RUNG wire#powerrail
      Contact( "Get Sinais de Interlock Main line".Station[9]."Sinal do job"[3] )
      Contact( "Get Sinais de Interlock Main line".Station[9]."Sinal do job"[4] )
      Contact( "Get Sinais de Interlock Main line".Station[9]."Sinal do job"[2] )
      Coil( "GAP_E_EIXO_PENDURADO" )
   END_RUNG
   // the same network as SCL:
   "GAP_E_EIXO_PENDURADO" := "Get Sinais de Interlock Main line".Station[9]."Sinal do job"[3] AND "Get Sinais de Interlock Main line".Station[9]."Sinal do job"[4] AND "Get Sinais de Interlock Main line".Station[9]."Sinal do job"[2];
END_REGION

REGION Network 38 (SCL): SEM JOB POKA YOKE P100 ORING MAP
   IF "EQUIPAMENTOS_RECIPE_POS_TAKT".EQUIPAMENTOS[17].RECIPE = 'ETRCALIP01' THEN
   "Put Sinais de Interlock Main line".RESERVED_4 := TRUE;
   ELSIF "BORDA_MD2".Q THEN
       "Put Sinais de Interlock Main line".RESERVED_4 := FALSE;
   END_IF;
END_REGION
END_FUNCTION
